ACTION act_Oper:
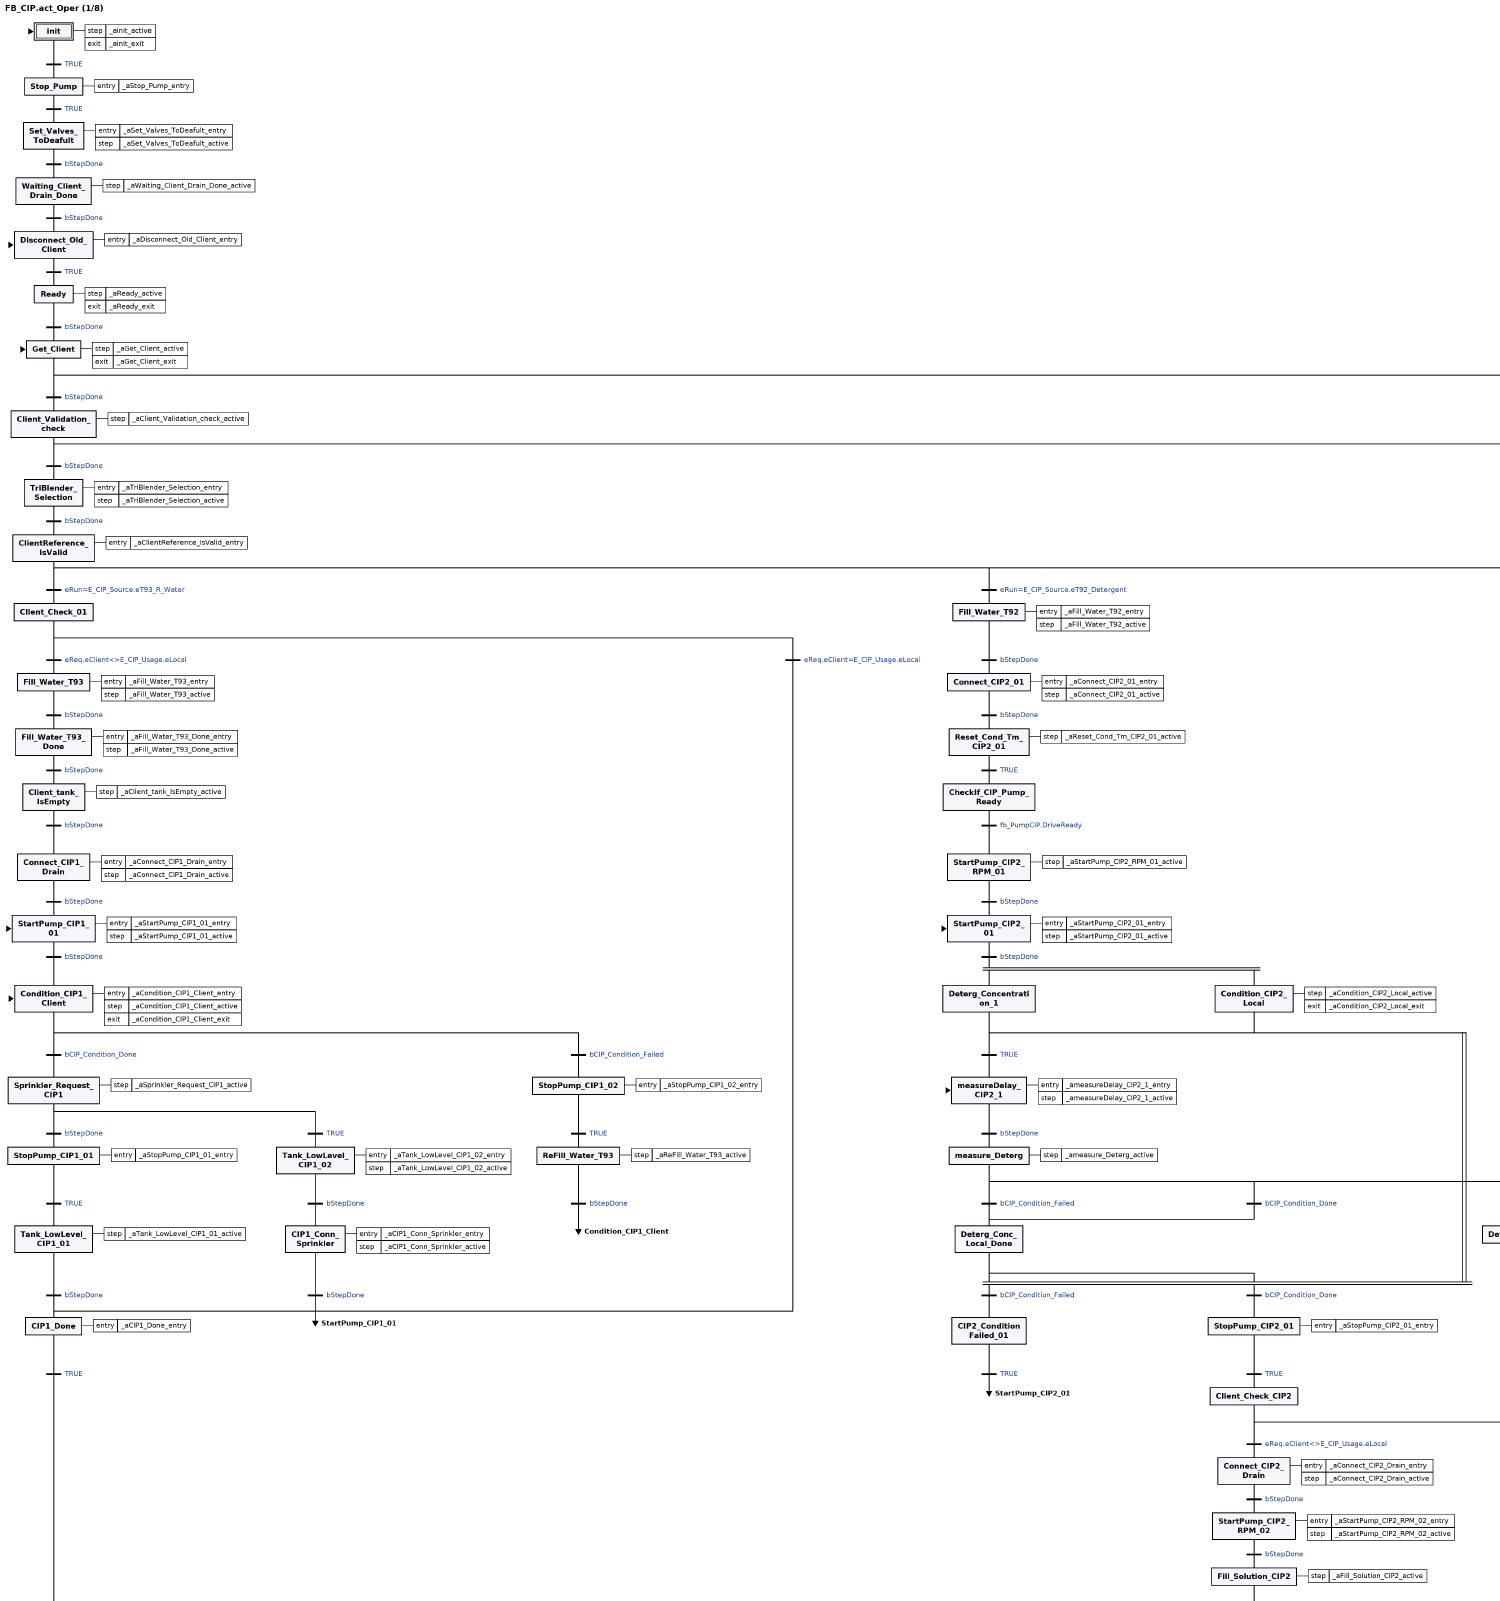
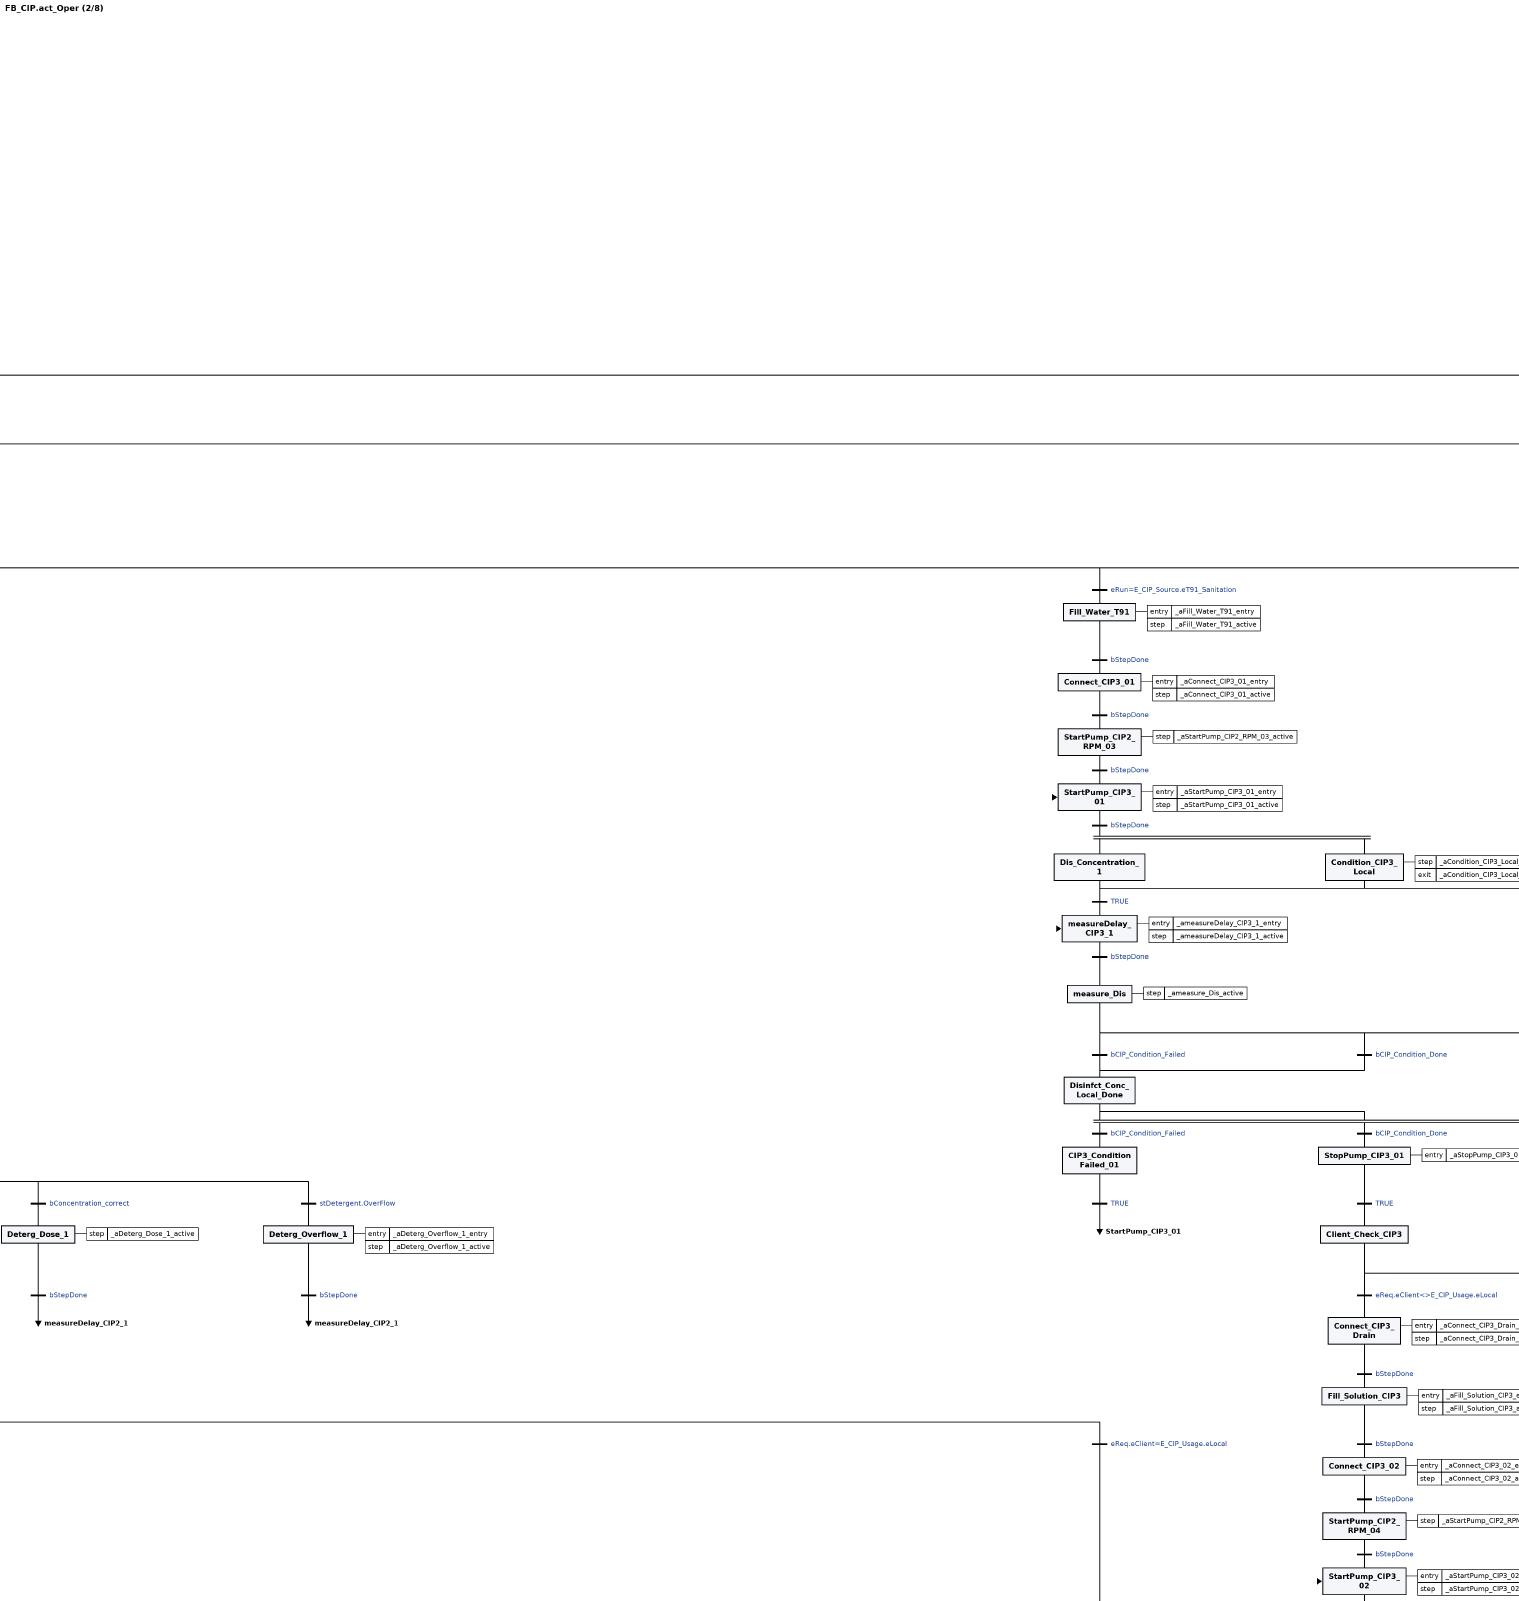
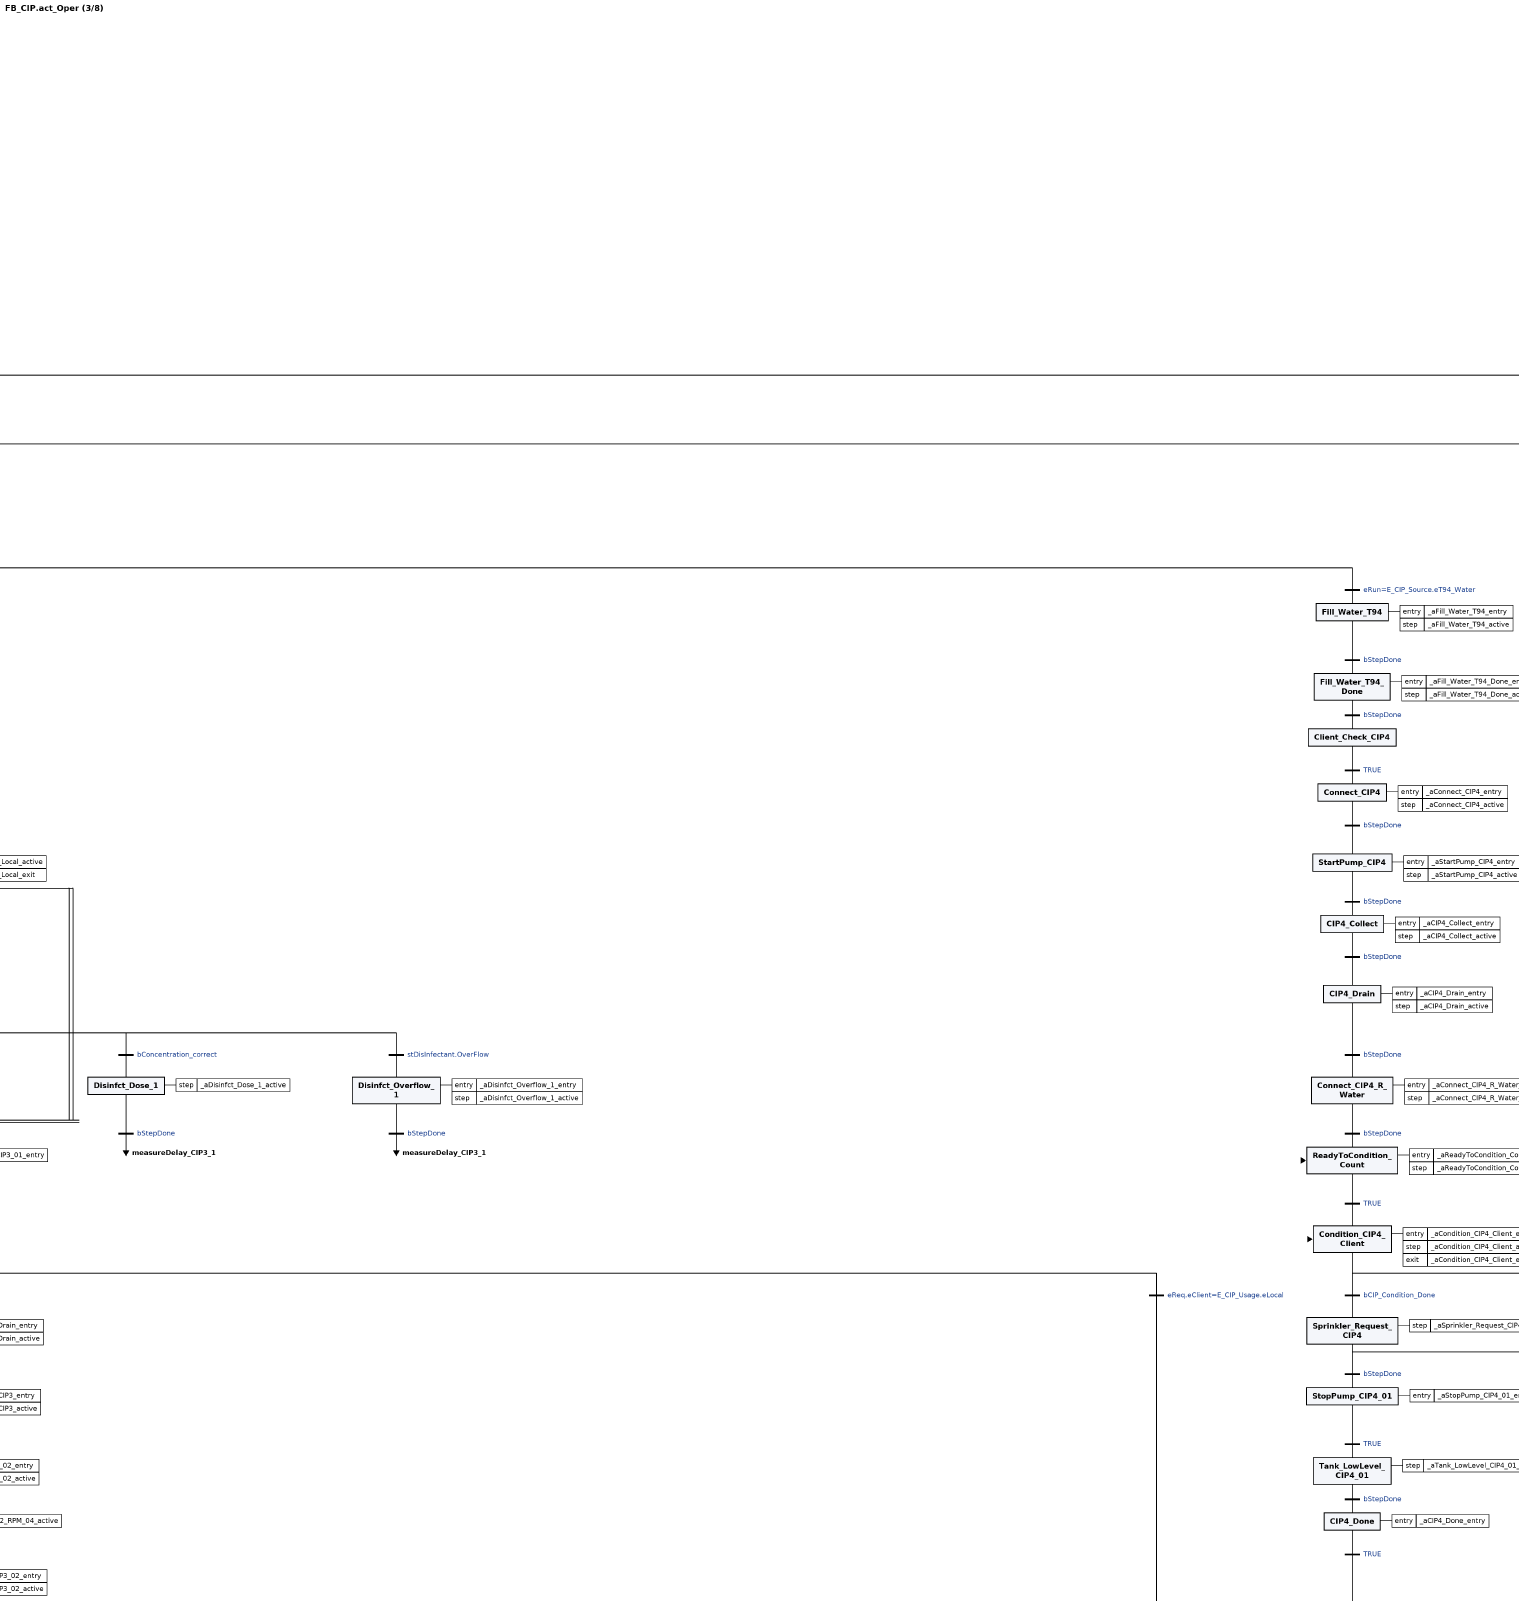
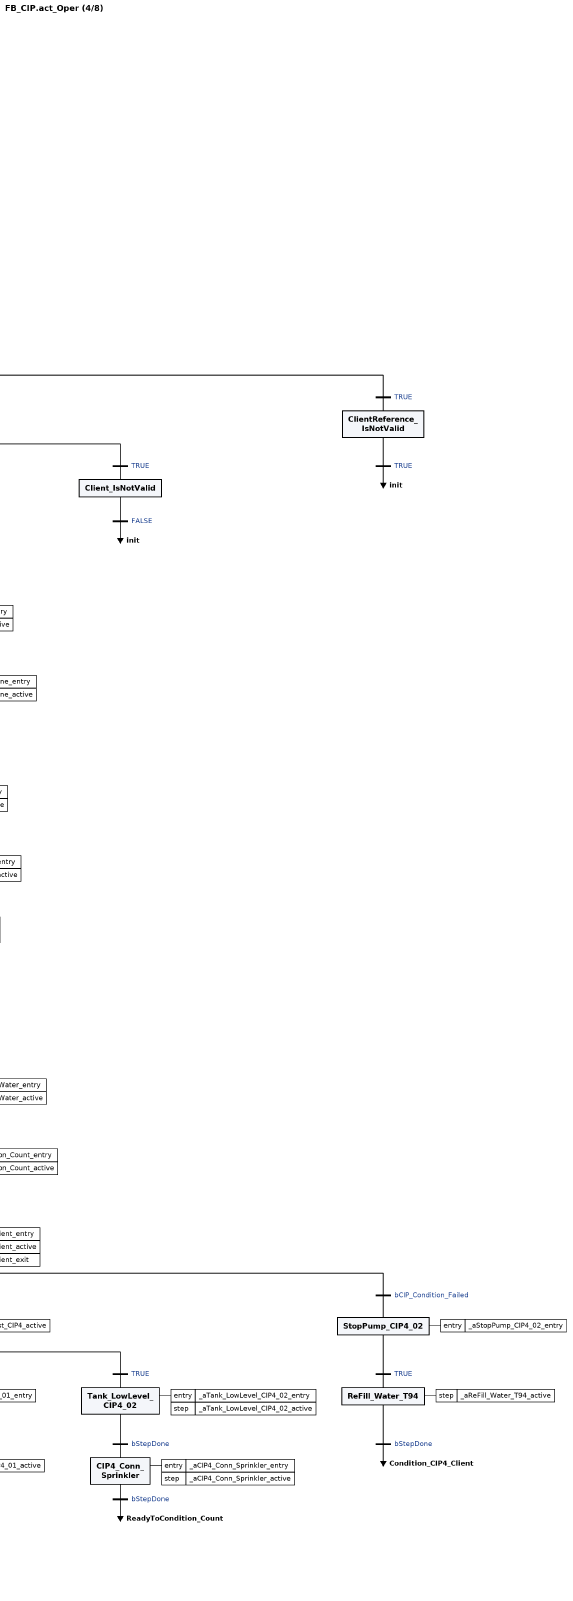
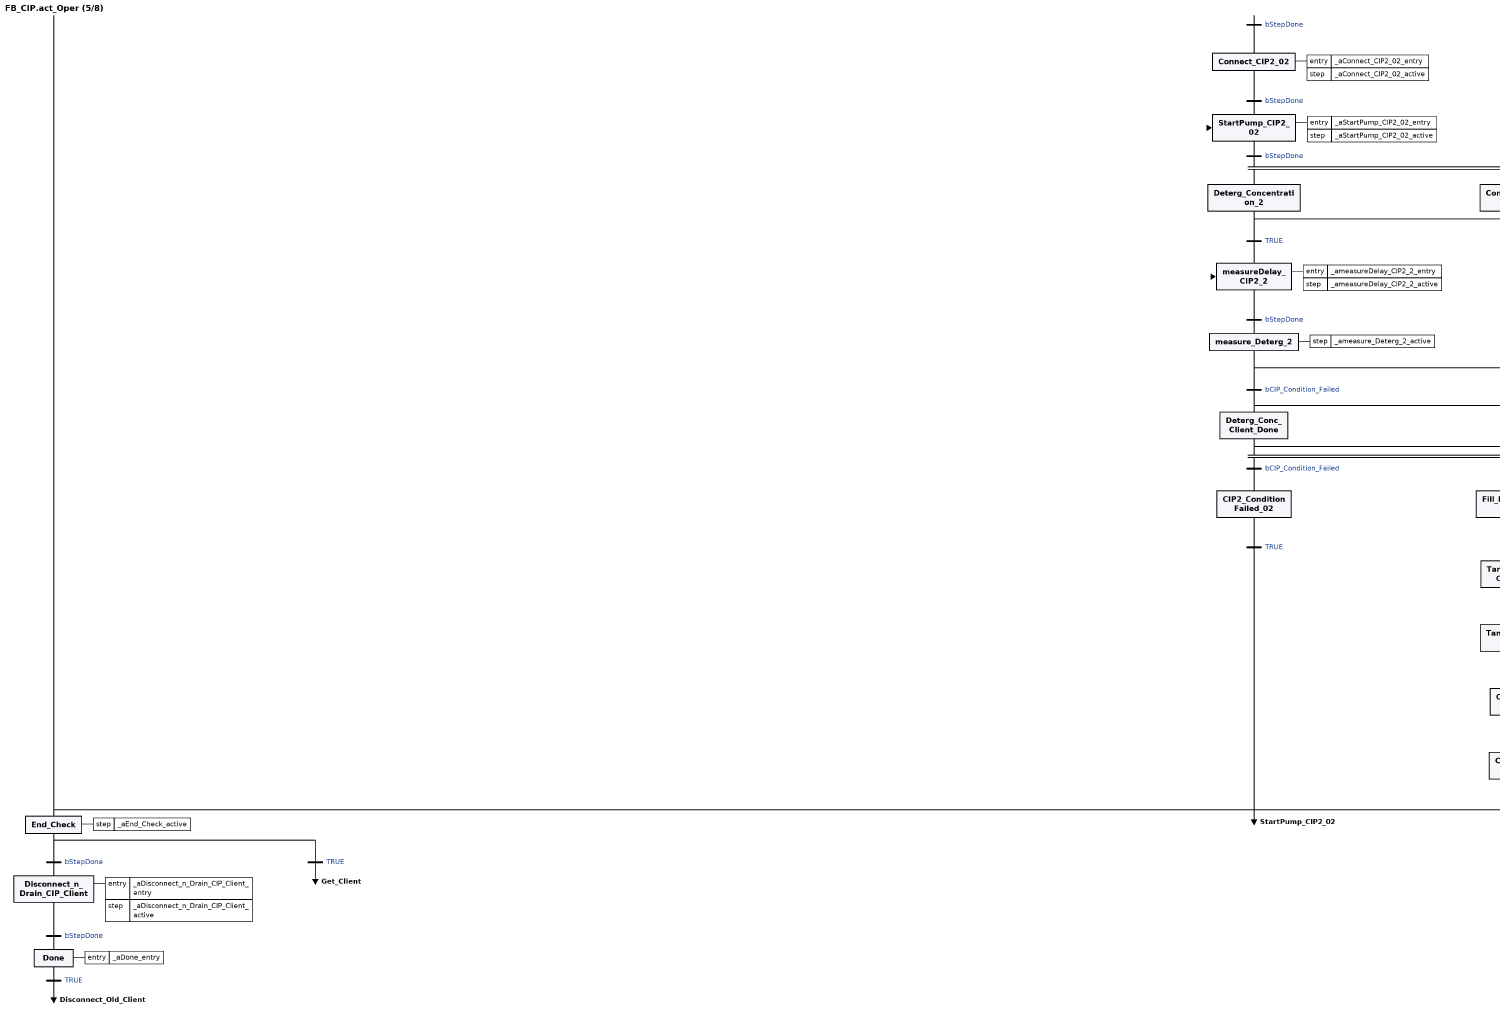
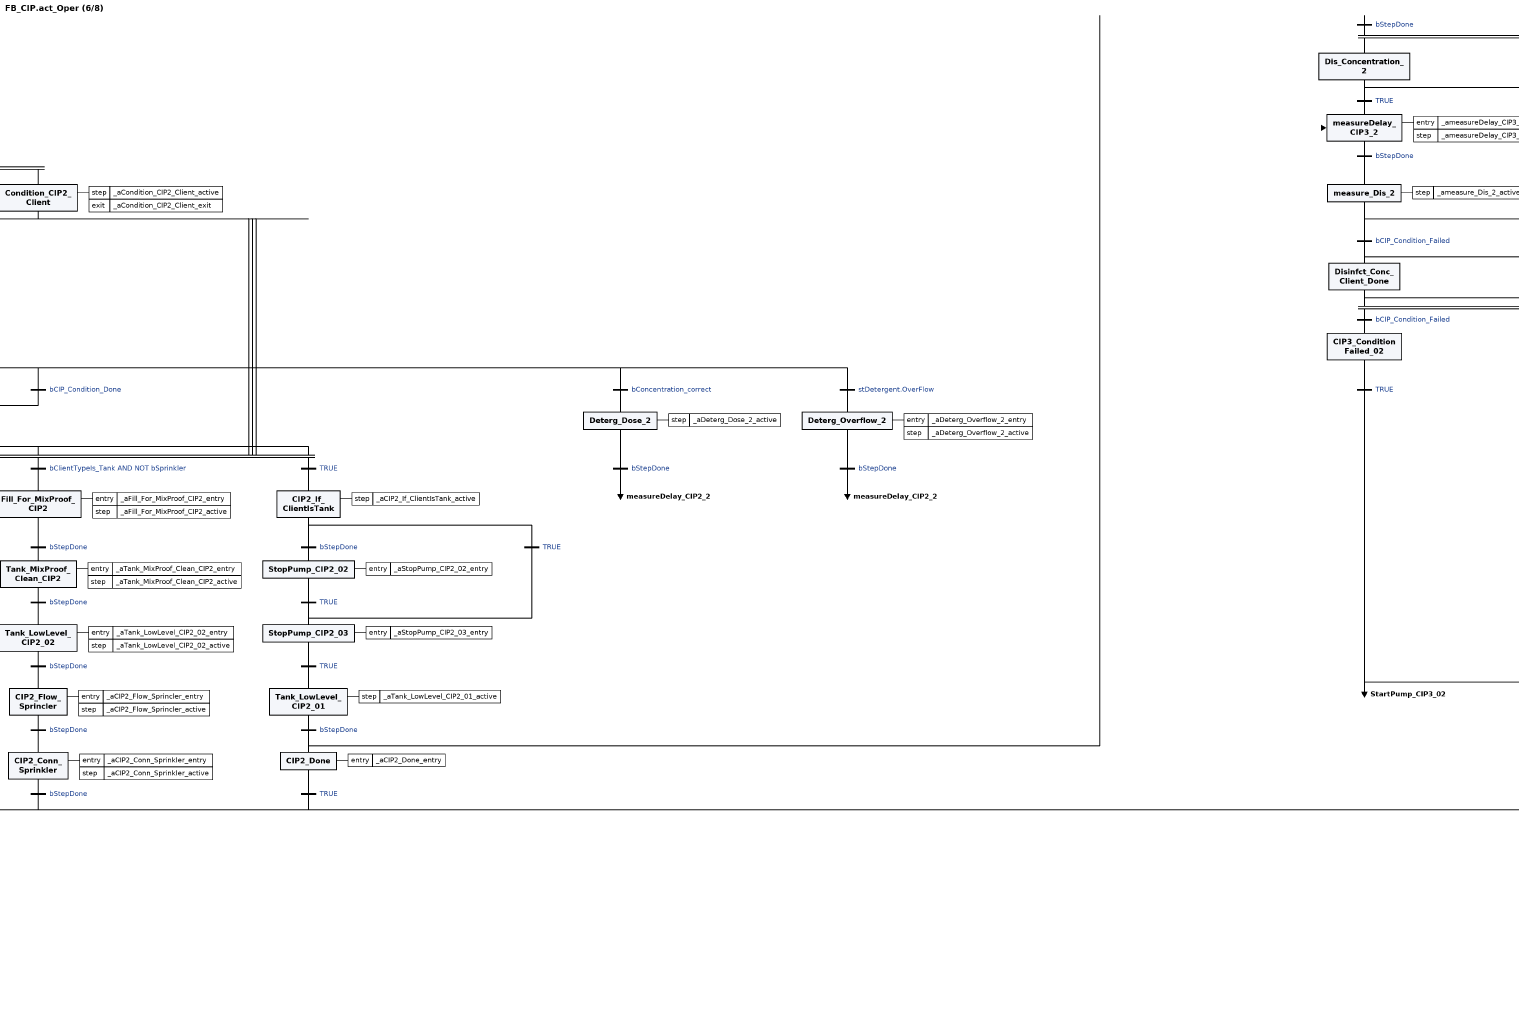
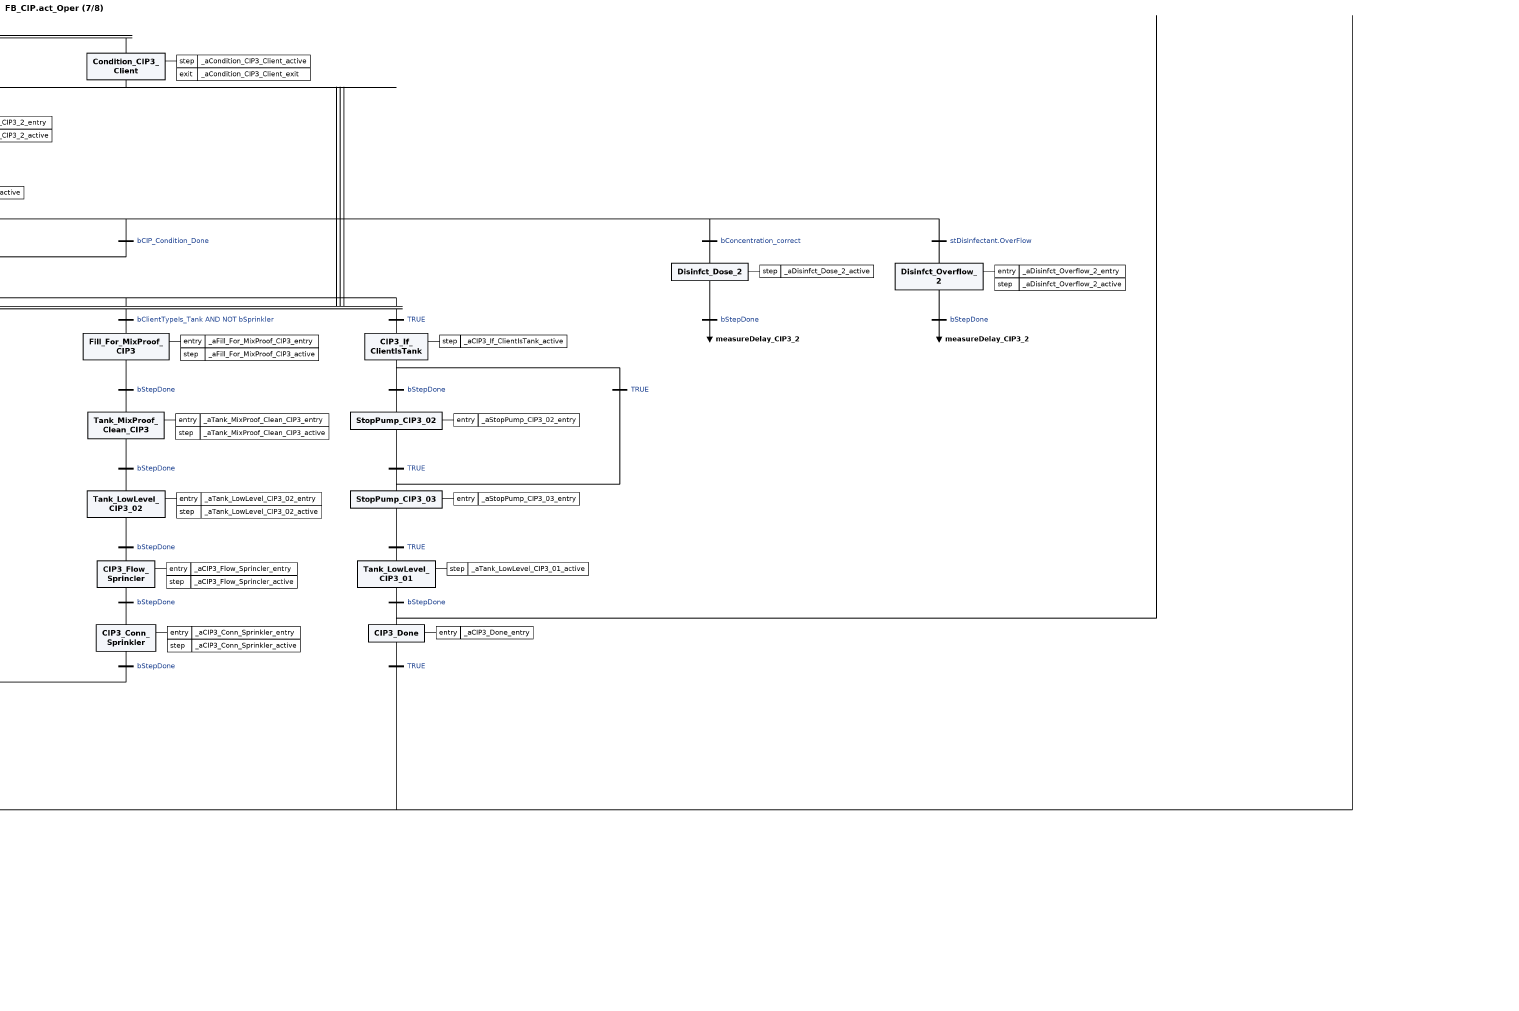
INITIAL_STEP init:
    _ainit_active(N);  // step action
    _ainit_exit(P0);  // exit action
END_STEP
TRANSITION FROM init TO Stop_Pump
    := TRUE;
END_TRANSITION
STEP Stop_Pump:
    _aStop_Pump_entry(P1);  // entry action
END_STEP
TRANSITION FROM Stop_Pump TO Set_Valves_ToDeafult
    := TRUE;
END_TRANSITION
STEP Set_Valves_ToDeafult:  // min time T#0.1s
    _aSet_Valves_ToDeafult_entry(P1);  // entry action
    _aSet_Valves_ToDeafult_active(N);  // step action
END_STEP
TRANSITION FROM Set_Valves_ToDeafult TO Waiting_Client_Drain_Done
    := bStepDone;
END_TRANSITION
STEP Waiting_Client_Drain_Done:  // min time T#0.1s
    _aWaiting_Client_Drain_Done_active(N);  // step action
END_STEP
TRANSITION FROM Waiting_Client_Drain_Done TO Disconnect_Old_Client
    := bStepDone;
END_TRANSITION
STEP Disconnect_Old_Client:
    _aDisconnect_Old_Client_entry(P1);  // entry action
END_STEP
TRANSITION FROM Disconnect_Old_Client TO Ready
    := TRUE;
END_TRANSITION
STEP Ready:
    _aReady_active(N);  // step action
    _aReady_exit(P0);  // exit action
END_STEP
TRANSITION FROM Ready TO Get_Client
    := bStepDone;
END_TRANSITION
STEP Get_Client:  // max time T#0.1s
    _aGet_Client_active(N);  // step action
    _aGet_Client_exit(P0);  // exit action
END_STEP
TRANSITION FROM Get_Client TO Client_Validation_check
    := bStepDone;
END_TRANSITION
TRANSITION FROM Get_Client TO ClientReference_IsNotValid
    := TRUE;
END_TRANSITION
STEP ClientReference_IsNotValid:  // min time T#2s
END_STEP
TRANSITION FROM ClientReference_IsNotValid TO init
    := TRUE;
END_TRANSITION
STEP Client_Validation_check:
    _aClient_Validation_check_active(N);  // step action
END_STEP
TRANSITION FROM Client_Validation_check TO TriBlender_Selection
    := bStepDone;
END_TRANSITION
STEP TriBlender_Selection:
    _aTriBlender_Selection_entry(P1);  // entry action
    _aTriBlender_Selection_active(N);  // step action
END_STEP
TRANSITION FROM TriBlender_Selection TO ClientReference_IsValid
    := bStepDone;
END_TRANSITION
TRANSITION FROM Client_Validation_check TO Client_IsNotValid
    := TRUE;
END_TRANSITION
STEP Client_IsNotValid:  // min time T#2s
END_STEP
TRANSITION FROM Client_IsNotValid TO init
    := FALSE;
END_TRANSITION
STEP ClientReference_IsValid:
    _aClientReference_IsValid_entry(P1);  // entry action
END_STEP
TRANSITION FROM ClientReference_IsValid TO Client_Check_01
    := eRun=E_CIP_Source.eT93_R_Water;
END_TRANSITION
// macro R_Water begins
STEP Client_Check_01:
END_STEP
TRANSITION FROM Client_Check_01 TO Fill_Water_T93
    := eReq.eClient<>E_CIP_Usage.eLocal;
END_TRANSITION
STEP Fill_Water_T93:
    _aFill_Water_T93_entry(P1);  // entry action
    _aFill_Water_T93_active(N);  // step action
END_STEP
TRANSITION FROM Fill_Water_T93 TO Fill_Water_T93_Done
    := bStepDone;
END_TRANSITION
STEP Fill_Water_T93_Done:
    _aFill_Water_T93_Done_entry(P1);  // entry action
    _aFill_Water_T93_Done_active(N);  // step action
END_STEP
TRANSITION FROM Fill_Water_T93_Done TO Client_tank_IsEmpty
    := bStepDone;
END_TRANSITION
STEP Client_tank_IsEmpty:  // min time T#5s
    _aClient_tank_IsEmpty_active(N);  // step action
END_STEP
TRANSITION FROM Client_tank_IsEmpty TO Connect_CIP1_Drain
    := bStepDone;
END_TRANSITION
STEP Connect_CIP1_Drain:
    _aConnect_CIP1_Drain_entry(P1);  // entry action
    _aConnect_CIP1_Drain_active(N);  // step action
END_STEP
TRANSITION FROM Connect_CIP1_Drain TO StartPump_CIP1_01
    := bStepDone;
END_TRANSITION
STEP StartPump_CIP1_01:
    _aStartPump_CIP1_01_entry(P1);  // entry action
    _aStartPump_CIP1_01_active(N);  // step action
END_STEP
TRANSITION FROM StartPump_CIP1_01 TO Condition_CIP1_Client
    := bStepDone;
END_TRANSITION
STEP Condition_CIP1_Client:
    _aCondition_CIP1_Client_entry(P1);  // entry action
    _aCondition_CIP1_Client_active(N);  // step action
    _aCondition_CIP1_Client_exit(P0);  // exit action
END_STEP
TRANSITION FROM Condition_CIP1_Client TO Sprinkler_Request_CIP1
    := bCIP_Condition_Done;
END_TRANSITION
STEP Sprinkler_Request_CIP1:
    _aSprinkler_Request_CIP1_active(N);  // step action
END_STEP
TRANSITION FROM Sprinkler_Request_CIP1 TO StopPump_CIP1_01
    := bStepDone;
END_TRANSITION
STEP StopPump_CIP1_01:
    _aStopPump_CIP1_01_entry(P1);  // entry action
END_STEP
TRANSITION FROM StopPump_CIP1_01 TO Tank_LowLevel_CIP1_01
    := TRUE;
END_TRANSITION
STEP Tank_LowLevel_CIP1_01:
    _aTank_LowLevel_CIP1_01_active(N);  // step action
END_STEP
TRANSITION FROM Tank_LowLevel_CIP1_01 TO CIP1_Done
    := bStepDone;
END_TRANSITION
TRANSITION FROM Sprinkler_Request_CIP1 TO Tank_LowLevel_CIP1_02
    := TRUE;
END_TRANSITION
STEP Tank_LowLevel_CIP1_02:
    _aTank_LowLevel_CIP1_02_entry(P1);  // entry action
    _aTank_LowLevel_CIP1_02_active(N);  // step action
END_STEP
TRANSITION FROM Tank_LowLevel_CIP1_02 TO CIP1_Conn_Sprinkler
    := bStepDone;
END_TRANSITION
STEP CIP1_Conn_Sprinkler:
    _aCIP1_Conn_Sprinkler_entry(P1);  // entry action
    _aCIP1_Conn_Sprinkler_active(N);  // step action
END_STEP
TRANSITION FROM CIP1_Conn_Sprinkler TO StartPump_CIP1_01
    := bStepDone;
END_TRANSITION
TRANSITION FROM Condition_CIP1_Client TO StopPump_CIP1_02
    := bCIP_Condition_Failed;
END_TRANSITION
STEP StopPump_CIP1_02:
    _aStopPump_CIP1_02_entry(P1);  // entry action
END_STEP
TRANSITION FROM StopPump_CIP1_02 TO ReFill_Water_T93
    := TRUE;
END_TRANSITION
STEP ReFill_Water_T93:
    _aReFill_Water_T93_active(N);  // step action
END_STEP
TRANSITION FROM ReFill_Water_T93 TO Condition_CIP1_Client
    := bStepDone;
END_TRANSITION
TRANSITION FROM Client_Check_01 TO CIP1_Done
    := eReq.eClient=E_CIP_Usage.eLocal;
END_TRANSITION
STEP CIP1_Done:  // min time T#2s
    _aCIP1_Done_entry(P1);  // entry action
END_STEP
TRANSITION FROM CIP1_Done TO End_Check
    := TRUE;
END_TRANSITION
TRANSITION FROM ClientReference_IsValid TO Fill_Water_T92
    := eRun=E_CIP_Source.eT92_Detergent;
END_TRANSITION
// macro Detergent begins
STEP Fill_Water_T92:
    _aFill_Water_T92_entry(P1);  // entry action
    _aFill_Water_T92_active(N);  // step action
END_STEP
TRANSITION FROM Fill_Water_T92 TO Connect_CIP2_01
    := bStepDone;
END_TRANSITION
STEP Connect_CIP2_01:
    _aConnect_CIP2_01_entry(P1);  // entry action
    _aConnect_CIP2_01_active(N);  // step action
END_STEP
TRANSITION FROM Connect_CIP2_01 TO Reset_Cond_Tm_CIP2_01
    := bStepDone;
END_TRANSITION
STEP Reset_Cond_Tm_CIP2_01:
    _aReset_Cond_Tm_CIP2_01_active(N);  // step action
END_STEP
TRANSITION FROM Reset_Cond_Tm_CIP2_01 TO CheckIf_CIP_Pump_Ready
    := TRUE;
END_TRANSITION
STEP CheckIf_CIP_Pump_Ready:
END_STEP
TRANSITION FROM CheckIf_CIP_Pump_Ready TO StartPump_CIP2_RPM_01
    := fb_PumpCIP.DriveReady;
END_TRANSITION
STEP StartPump_CIP2_RPM_01:
    _aStartPump_CIP2_RPM_01_active(N);  // step action
END_STEP
TRANSITION FROM StartPump_CIP2_RPM_01 TO StartPump_CIP2_01
    := bStepDone;
END_TRANSITION
STEP StartPump_CIP2_01:  // min time T#2s
    _aStartPump_CIP2_01_entry(P1);  // entry action
    _aStartPump_CIP2_01_active(N);  // step action
END_STEP
TRANSITION FROM StartPump_CIP2_01 TO (Deterg_Concentration_1, Condition_CIP2_Local)
    := bStepDone;
END_TRANSITION
STEP Deterg_Concentration_1:
END_STEP
TRANSITION FROM Deterg_Concentration_1 TO measureDelay_CIP2_1
    := TRUE;
END_TRANSITION
STEP measureDelay_CIP2_1:
    _ameasureDelay_CIP2_1_entry(P1);  // entry action
    _ameasureDelay_CIP2_1_active(N);  // step action
END_STEP
TRANSITION FROM measureDelay_CIP2_1 TO measure_Deterg
    := bStepDone;
END_TRANSITION
STEP measure_Deterg:  // min time t#1s
    _ameasure_Deterg_active(N);  // step action
END_STEP
TRANSITION FROM measure_Deterg TO Deterg_Conc_Local_Done
    := bCIP_Condition_Failed;
END_TRANSITION
TRANSITION FROM measure_Deterg TO Deterg_Conc_Local_Done
    := bCIP_Condition_Done;
END_TRANSITION
TRANSITION FROM measure_Deterg TO Deterg_Dose_1
    := bConcentration_correct;
END_TRANSITION
STEP Deterg_Dose_1:
    _aDeterg_Dose_1_active(N);  // step action
END_STEP
TRANSITION FROM Deterg_Dose_1 TO measureDelay_CIP2_1
    := bStepDone;
END_TRANSITION
TRANSITION FROM measure_Deterg TO Deterg_Overflow_1
    := stDetergent.OverFlow;
END_TRANSITION
STEP Deterg_Overflow_1:
    _aDeterg_Overflow_1_entry(P1);  // entry action
    _aDeterg_Overflow_1_active(N);  // step action
END_STEP
TRANSITION FROM Deterg_Overflow_1 TO measureDelay_CIP2_1
    := bStepDone;
END_TRANSITION
STEP Deterg_Conc_Local_Done:
END_STEP
STEP Condition_CIP2_Local:
    _aCondition_CIP2_Local_active(N);  // step action
    _aCondition_CIP2_Local_exit(P0);  // exit action
END_STEP
TRANSITION FROM (Deterg_Conc_Local_Done, Condition_CIP2_Local) TO CIP2_ConditionFailed_01
    := bCIP_Condition_Failed;
END_TRANSITION
STEP CIP2_ConditionFailed_01:
END_STEP
TRANSITION FROM CIP2_ConditionFailed_01 TO StartPump_CIP2_01
    := TRUE;
END_TRANSITION
TRANSITION FROM (Deterg_Conc_Local_Done, Condition_CIP2_Local) TO StopPump_CIP2_01
    := bCIP_Condition_Done;
END_TRANSITION
STEP StopPump_CIP2_01:
    _aStopPump_CIP2_01_entry(P1);  // entry action
END_STEP
TRANSITION FROM StopPump_CIP2_01 TO Client_Check_CIP2
    := TRUE;
END_TRANSITION
STEP Client_Check_CIP2:
END_STEP
TRANSITION FROM Client_Check_CIP2 TO Connect_CIP2_Drain
    := eReq.eClient<>E_CIP_Usage.eLocal;
END_TRANSITION
STEP Connect_CIP2_Drain:
    _aConnect_CIP2_Drain_entry(P1);  // entry action
    _aConnect_CIP2_Drain_active(N);  // step action
END_STEP
TRANSITION FROM Connect_CIP2_Drain TO StartPump_CIP2_RPM_02
    := bStepDone;
END_TRANSITION
STEP StartPump_CIP2_RPM_02:
    _aStartPump_CIP2_RPM_02_entry(P1);  // entry action
    _aStartPump_CIP2_RPM_02_active(N);  // step action
END_STEP
TRANSITION FROM StartPump_CIP2_RPM_02 TO Fill_Solution_CIP2
    := bStepDone;
END_TRANSITION
STEP Fill_Solution_CIP2:
    _aFill_Solution_CIP2_active(N);  // step action
END_STEP
TRANSITION FROM Fill_Solution_CIP2 TO Connect_CIP2_02
    := bStepDone;
END_TRANSITION
STEP Connect_CIP2_02:
    _aConnect_CIP2_02_entry(P1);  // entry action
    _aConnect_CIP2_02_active(N);  // step action
END_STEP
TRANSITION FROM Connect_CIP2_02 TO StartPump_CIP2_02
    := bStepDone;
END_TRANSITION
STEP StartPump_CIP2_02:  // min time T#2s
    _aStartPump_CIP2_02_entry(P1);  // entry action
    _aStartPump_CIP2_02_active(N);  // step action
END_STEP
TRANSITION FROM StartPump_CIP2_02 TO (Deterg_Concentration_2, Condition_CIP2_Client)
    := bStepDone;
END_TRANSITION
STEP Deterg_Concentration_2:
END_STEP
TRANSITION FROM Deterg_Concentration_2 TO measureDelay_CIP2_2
    := TRUE;
END_TRANSITION
STEP measureDelay_CIP2_2:
    _ameasureDelay_CIP2_2_entry(P1);  // entry action
    _ameasureDelay_CIP2_2_active(N);  // step action
END_STEP
TRANSITION FROM measureDelay_CIP2_2 TO measure_Deterg_2
    := bStepDone;
END_TRANSITION
STEP measure_Deterg_2:  // min time t#1s
    _ameasure_Deterg_2_active(N);  // step action
END_STEP
TRANSITION FROM measure_Deterg_2 TO Deterg_Conc_Client_Done
    := bCIP_Condition_Failed;
END_TRANSITION
TRANSITION FROM measure_Deterg_2 TO Deterg_Conc_Client_Done
    := bCIP_Condition_Done;
END_TRANSITION
TRANSITION FROM measure_Deterg_2 TO Deterg_Dose_2
    := bConcentration_correct;
END_TRANSITION
STEP Deterg_Dose_2:
    _aDeterg_Dose_2_active(N);  // step action
END_STEP
TRANSITION FROM Deterg_Dose_2 TO measureDelay_CIP2_2
    := bStepDone;
END_TRANSITION
TRANSITION FROM measure_Deterg_2 TO Deterg_Overflow_2
    := stDetergent.OverFlow;
END_TRANSITION
STEP Deterg_Overflow_2:
    _aDeterg_Overflow_2_entry(P1);  // entry action
    _aDeterg_Overflow_2_active(N);  // step action
END_STEP
TRANSITION FROM Deterg_Overflow_2 TO measureDelay_CIP2_2
    := bStepDone;
END_TRANSITION
STEP Deterg_Conc_Client_Done:
END_STEP
STEP Condition_CIP2_Client:
    _aCondition_CIP2_Client_active(N);  // step action
    _aCondition_CIP2_Client_exit(P0);  // exit action
END_STEP
TRANSITION FROM (Deterg_Conc_Client_Done, Condition_CIP2_Client) TO CIP2_ConditionFailed_02
    := bCIP_Condition_Failed;
END_TRANSITION
STEP CIP2_ConditionFailed_02:
END_STEP
TRANSITION FROM CIP2_ConditionFailed_02 TO StartPump_CIP2_02
    := TRUE;
END_TRANSITION
TRANSITION FROM (Deterg_Conc_Client_Done, Condition_CIP2_Client) TO Fill_For_MixProof_CIP2
    := bClientTypeIs_Tank AND NOT bSprinkler;
END_TRANSITION
STEP Fill_For_MixProof_CIP2:
    _aFill_For_MixProof_CIP2_entry(P1);  // entry action
    _aFill_For_MixProof_CIP2_active(N);  // step action
END_STEP
TRANSITION FROM Fill_For_MixProof_CIP2 TO Tank_MixProof_Clean_CIP2
    := bStepDone;
END_TRANSITION
STEP Tank_MixProof_Clean_CIP2:
    _aTank_MixProof_Clean_CIP2_entry(P1);  // entry action
    _aTank_MixProof_Clean_CIP2_active(N);  // step action
END_STEP
TRANSITION FROM Tank_MixProof_Clean_CIP2 TO Tank_LowLevel_CIP2_02
    := bStepDone;
END_TRANSITION
STEP Tank_LowLevel_CIP2_02:
    _aTank_LowLevel_CIP2_02_entry(P1);  // entry action
    _aTank_LowLevel_CIP2_02_active(N);  // step action
END_STEP
TRANSITION FROM Tank_LowLevel_CIP2_02 TO CIP2_Flow_Sprincler
    := bStepDone;
END_TRANSITION
STEP CIP2_Flow_Sprincler:
    _aCIP2_Flow_Sprincler_entry(P1);  // entry action
    _aCIP2_Flow_Sprincler_active(N);  // step action
END_STEP
TRANSITION FROM CIP2_Flow_Sprincler TO CIP2_Conn_Sprinkler
    := bStepDone;
END_TRANSITION
STEP CIP2_Conn_Sprinkler:
    _aCIP2_Conn_Sprinkler_entry(P1);  // entry action
    _aCIP2_Conn_Sprinkler_active(N);  // step action
END_STEP
TRANSITION FROM CIP2_Conn_Sprinkler TO StartPump_CIP2_02
    := bStepDone;
END_TRANSITION
TRANSITION FROM (Deterg_Conc_Client_Done, Condition_CIP2_Client) TO CIP2_If_ClientIsTank
    := TRUE;
END_TRANSITION
STEP CIP2_If_ClientIsTank:
    _aCIP2_If_ClientIsTank_active(N);  // step action
END_STEP
TRANSITION FROM CIP2_If_ClientIsTank TO StopPump_CIP2_02
    := bStepDone;
END_TRANSITION
STEP StopPump_CIP2_02:
    _aStopPump_CIP2_02_entry(P1);  // entry action
END_STEP
TRANSITION FROM StopPump_CIP2_02 TO StopPump_CIP2_03
    := TRUE;
END_TRANSITION
TRANSITION FROM CIP2_If_ClientIsTank TO StopPump_CIP2_03
    := TRUE;
END_TRANSITION
STEP StopPump_CIP2_03:
    _aStopPump_CIP2_03_entry(P1);  // entry action
END_STEP
TRANSITION FROM StopPump_CIP2_03 TO Tank_LowLevel_CIP2_01
    := TRUE;
END_TRANSITION
STEP Tank_LowLevel_CIP2_01:
    _aTank_LowLevel_CIP2_01_active(N);  // step action
END_STEP
TRANSITION FROM Tank_LowLevel_CIP2_01 TO CIP2_Done
    := bStepDone;
END_TRANSITION
TRANSITION FROM Client_Check_CIP2 TO CIP2_Done
    := eReq.eClient=E_CIP_Usage.eLocal;
END_TRANSITION
STEP CIP2_Done:  // min time T#2s
    _aCIP2_Done_entry(P1);  // entry action
END_STEP
TRANSITION FROM CIP2_Done TO End_Check
    := TRUE;
END_TRANSITION
TRANSITION FROM ClientReference_IsValid TO Fill_Water_T91
    := eRun=E_CIP_Source.eT91_Sanitation;
END_TRANSITION
// macro DisInfection begins
STEP Fill_Water_T91:
    _aFill_Water_T91_entry(P1);  // entry action
    _aFill_Water_T91_active(N);  // step action
END_STEP
TRANSITION FROM Fill_Water_T91 TO Connect_CIP3_01
    := bStepDone;
END_TRANSITION
STEP Connect_CIP3_01:
    _aConnect_CIP3_01_entry(P1);  // entry action
    _aConnect_CIP3_01_active(N);  // step action
END_STEP
TRANSITION FROM Connect_CIP3_01 TO StartPump_CIP2_RPM_03
    := bStepDone;
END_TRANSITION
STEP StartPump_CIP2_RPM_03:
    _aStartPump_CIP2_RPM_03_active(N);  // step action
END_STEP
TRANSITION FROM StartPump_CIP2_RPM_03 TO StartPump_CIP3_01
    := bStepDone;
END_TRANSITION
STEP StartPump_CIP3_01:  // min time T#3s
    _aStartPump_CIP3_01_entry(P1);  // entry action
    _aStartPump_CIP3_01_active(N);  // step action
END_STEP
TRANSITION FROM StartPump_CIP3_01 TO (Dis_Concentration_1, Condition_CIP3_Local)
    := bStepDone;
END_TRANSITION
STEP Dis_Concentration_1:
END_STEP
TRANSITION FROM Dis_Concentration_1 TO measureDelay_CIP3_1
    := TRUE;
END_TRANSITION
STEP measureDelay_CIP3_1:
    _ameasureDelay_CIP3_1_entry(P1);  // entry action
    _ameasureDelay_CIP3_1_active(N);  // step action
END_STEP
TRANSITION FROM measureDelay_CIP3_1 TO measure_Dis
    := bStepDone;
END_TRANSITION
STEP measure_Dis:  // min time t#1s
    _ameasure_Dis_active(N);  // step action
END_STEP
TRANSITION FROM measure_Dis TO Disinfct_Conc_Local_Done
    := bCIP_Condition_Failed;
END_TRANSITION
TRANSITION FROM measure_Dis TO Disinfct_Conc_Local_Done
    := bCIP_Condition_Done;
END_TRANSITION
TRANSITION FROM measure_Dis TO Disinfct_Dose_1
    := bConcentration_correct;
END_TRANSITION
STEP Disinfct_Dose_1:
    _aDisinfct_Dose_1_active(N);  // step action
END_STEP
TRANSITION FROM Disinfct_Dose_1 TO measureDelay_CIP3_1
    := bStepDone;
END_TRANSITION
TRANSITION FROM measure_Dis TO Disinfct_Overflow_1
    := stDisInfectant.OverFlow;
END_TRANSITION
STEP Disinfct_Overflow_1:
    _aDisinfct_Overflow_1_entry(P1);  // entry action
    _aDisinfct_Overflow_1_active(N);  // step action
END_STEP
TRANSITION FROM Disinfct_Overflow_1 TO measureDelay_CIP3_1
    := bStepDone;
END_TRANSITION
STEP Disinfct_Conc_Local_Done:
END_STEP
STEP Condition_CIP3_Local:
    _aCondition_CIP3_Local_active(N);  // step action
    _aCondition_CIP3_Local_exit(P0);  // exit action
END_STEP
TRANSITION FROM (Disinfct_Conc_Local_Done, Condition_CIP3_Local) TO CIP3_ConditionFailed_01
    := bCIP_Condition_Failed;
END_TRANSITION
STEP CIP3_ConditionFailed_01:
END_STEP
TRANSITION FROM CIP3_ConditionFailed_01 TO StartPump_CIP3_01
    := TRUE;
END_TRANSITION
TRANSITION FROM (Disinfct_Conc_Local_Done, Condition_CIP3_Local) TO StopPump_CIP3_01
    := bCIP_Condition_Done;
END_TRANSITION
STEP StopPump_CIP3_01:  // min time T#5s
    _aStopPump_CIP3_01_entry(P1);  // entry action
END_STEP
TRANSITION FROM StopPump_CIP3_01 TO Client_Check_CIP3
    := TRUE;
END_TRANSITION
STEP Client_Check_CIP3:
END_STEP
TRANSITION FROM Client_Check_CIP3 TO Connect_CIP3_Drain
    := eReq.eClient<>E_CIP_Usage.eLocal;
END_TRANSITION
STEP Connect_CIP3_Drain:
    _aConnect_CIP3_Drain_entry(P1);  // entry action
    _aConnect_CIP3_Drain_active(N);  // step action
END_STEP
TRANSITION FROM Connect_CIP3_Drain TO Fill_Solution_CIP3
    := bStepDone;
END_TRANSITION
STEP Fill_Solution_CIP3:
    _aFill_Solution_CIP3_entry(P1);  // entry action
    _aFill_Solution_CIP3_active(N);  // step action
END_STEP
TRANSITION FROM Fill_Solution_CIP3 TO Connect_CIP3_02
    := bStepDone;
END_TRANSITION
STEP Connect_CIP3_02:
    _aConnect_CIP3_02_entry(P1);  // entry action
    _aConnect_CIP3_02_active(N);  // step action
END_STEP
TRANSITION FROM Connect_CIP3_02 TO StartPump_CIP2_RPM_04
    := bStepDone;
END_TRANSITION
STEP StartPump_CIP2_RPM_04:
    _aStartPump_CIP2_RPM_04_active(N);  // step action
END_STEP
TRANSITION FROM StartPump_CIP2_RPM_04 TO StartPump_CIP3_02
    := bStepDone;
END_TRANSITION
STEP StartPump_CIP3_02:  // min time T#1s
    _aStartPump_CIP3_02_entry(P1);  // entry action
    _aStartPump_CIP3_02_active(N);  // step action
END_STEP
TRANSITION FROM StartPump_CIP3_02 TO (Dis_Concentration_2, Condition_CIP3_Client)
    := bStepDone;
END_TRANSITION
STEP Dis_Concentration_2:
END_STEP
TRANSITION FROM Dis_Concentration_2 TO measureDelay_CIP3_2
    := TRUE;
END_TRANSITION
STEP measureDelay_CIP3_2:
    _ameasureDelay_CIP3_2_entry(P1);  // entry action
    _ameasureDelay_CIP3_2_active(N);  // step action
END_STEP
TRANSITION FROM measureDelay_CIP3_2 TO measure_Dis_2
    := bStepDone;
END_TRANSITION
STEP measure_Dis_2:  // min time t#1s
    _ameasure_Dis_2_active(N);  // step action
END_STEP
TRANSITION FROM measure_Dis_2 TO Disinfct_Conc_Client_Done
    := bCIP_Condition_Failed;
END_TRANSITION
TRANSITION FROM measure_Dis_2 TO Disinfct_Conc_Client_Done
    := bCIP_Condition_Done;
END_TRANSITION
TRANSITION FROM measure_Dis_2 TO Disinfct_Dose_2
    := bConcentration_correct;
END_TRANSITION
STEP Disinfct_Dose_2:
    _aDisinfct_Dose_2_active(N);  // step action
END_STEP
TRANSITION FROM Disinfct_Dose_2 TO measureDelay_CIP3_2
    := bStepDone;
END_TRANSITION
TRANSITION FROM measure_Dis_2 TO Disinfct_Overflow_2
    := stDisInfectant.OverFlow;
END_TRANSITION
STEP Disinfct_Overflow_2:
    _aDisinfct_Overflow_2_entry(P1);  // entry action
    _aDisinfct_Overflow_2_active(N);  // step action
END_STEP
TRANSITION FROM Disinfct_Overflow_2 TO measureDelay_CIP3_2
    := bStepDone;
END_TRANSITION
STEP Disinfct_Conc_Client_Done:
END_STEP
STEP Condition_CIP3_Client:
    _aCondition_CIP3_Client_active(N);  // step action
    _aCondition_CIP3_Client_exit(P0);  // exit action
END_STEP
TRANSITION FROM (Disinfct_Conc_Client_Done, Condition_CIP3_Client) TO CIP3_ConditionFailed_02
    := bCIP_Condition_Failed;
END_TRANSITION
STEP CIP3_ConditionFailed_02:
END_STEP
TRANSITION FROM CIP3_ConditionFailed_02 TO StartPump_CIP3_02
    := TRUE;
END_TRANSITION
TRANSITION FROM (Disinfct_Conc_Client_Done, Condition_CIP3_Client) TO Fill_For_MixProof_CIP3
    := bClientTypeIs_Tank AND NOT bSprinkler;
END_TRANSITION
STEP Fill_For_MixProof_CIP3:
    _aFill_For_MixProof_CIP3_entry(P1);  // entry action
    _aFill_For_MixProof_CIP3_active(N);  // step action
END_STEP
TRANSITION FROM Fill_For_MixProof_CIP3 TO Tank_MixProof_Clean_CIP3
    := bStepDone;
END_TRANSITION
STEP Tank_MixProof_Clean_CIP3:
    _aTank_MixProof_Clean_CIP3_entry(P1);  // entry action
    _aTank_MixProof_Clean_CIP3_active(N);  // step action
END_STEP
TRANSITION FROM Tank_MixProof_Clean_CIP3 TO Tank_LowLevel_CIP3_02
    := bStepDone;
END_TRANSITION
STEP Tank_LowLevel_CIP3_02:
    _aTank_LowLevel_CIP3_02_entry(P1);  // entry action
    _aTank_LowLevel_CIP3_02_active(N);  // step action
END_STEP
TRANSITION FROM Tank_LowLevel_CIP3_02 TO CIP3_Flow_Sprincler
    := bStepDone;
END_TRANSITION
STEP CIP3_Flow_Sprincler:
    _aCIP3_Flow_Sprincler_entry(P1);  // entry action
    _aCIP3_Flow_Sprincler_active(N);  // step action
END_STEP
TRANSITION FROM CIP3_Flow_Sprincler TO CIP3_Conn_Sprinkler
    := bStepDone;
END_TRANSITION
STEP CIP3_Conn_Sprinkler:
    _aCIP3_Conn_Sprinkler_entry(P1);  // entry action
    _aCIP3_Conn_Sprinkler_active(N);  // step action
END_STEP
TRANSITION FROM CIP3_Conn_Sprinkler TO StartPump_CIP3_02
    := bStepDone;
END_TRANSITION
TRANSITION FROM (Disinfct_Conc_Client_Done, Condition_CIP3_Client) TO CIP3_If_ClientIsTank
    := TRUE;
END_TRANSITION
STEP CIP3_If_ClientIsTank:
    _aCIP3_If_ClientIsTank_active(N);  // step action
END_STEP
TRANSITION FROM CIP3_If_ClientIsTank TO StopPump_CIP3_02
    := bStepDone;
END_TRANSITION
STEP StopPump_CIP3_02:  // min time T#2s
    _aStopPump_CIP3_02_entry(P1);  // entry action
END_STEP
TRANSITION FROM StopPump_CIP3_02 TO StopPump_CIP3_03
    := TRUE;
END_TRANSITION
TRANSITION FROM CIP3_If_ClientIsTank TO StopPump_CIP3_03
    := TRUE;
END_TRANSITION
STEP StopPump_CIP3_03:
    _aStopPump_CIP3_03_entry(P1);  // entry action
END_STEP
TRANSITION FROM StopPump_CIP3_03 TO Tank_LowLevel_CIP3_01
    := TRUE;
END_TRANSITION
STEP Tank_LowLevel_CIP3_01:
    _aTank_LowLevel_CIP3_01_active(N);  // step action
END_STEP
TRANSITION FROM Tank_LowLevel_CIP3_01 TO CIP3_Done
    := bStepDone;
END_TRANSITION
TRANSITION FROM Client_Check_CIP3 TO CIP3_Done
    := eReq.eClient=E_CIP_Usage.eLocal;
END_TRANSITION
STEP CIP3_Done:  // min time T#2s
    _aCIP3_Done_entry(P1);  // entry action
END_STEP
TRANSITION FROM CIP3_Done TO End_Check
    := TRUE;
END_TRANSITION
TRANSITION FROM ClientReference_IsValid TO Fill_Water_T94
    := eRun=E_CIP_Source.eT94_Water;
END_TRANSITION
// macro Water begins
STEP Fill_Water_T94:
    _aFill_Water_T94_entry(P1);  // entry action
    _aFill_Water_T94_active(N);  // step action
END_STEP
TRANSITION FROM Fill_Water_T94 TO Fill_Water_T94_Done
    := bStepDone;
END_TRANSITION
STEP Fill_Water_T94_Done:
    _aFill_Water_T94_Done_entry(P1);  // entry action
    _aFill_Water_T94_Done_active(N);  // step action
END_STEP
TRANSITION FROM Fill_Water_T94_Done TO Client_Check_CIP4
    := bStepDone;
END_TRANSITION
STEP Client_Check_CIP4:
END_STEP
TRANSITION FROM Client_Check_CIP4 TO Connect_CIP4
    := TRUE;
END_TRANSITION
STEP Connect_CIP4:
    _aConnect_CIP4_entry(P1);  // entry action
    _aConnect_CIP4_active(N);  // step action
END_STEP
TRANSITION FROM Connect_CIP4 TO StartPump_CIP4
    := bStepDone;
END_TRANSITION
STEP StartPump_CIP4:  // min time T#3s
    _aStartPump_CIP4_entry(P1);  // entry action
    _aStartPump_CIP4_active(N);  // step action
END_STEP
TRANSITION FROM StartPump_CIP4 TO CIP4_Collect
    := bStepDone;
END_TRANSITION
STEP CIP4_Collect:  // min time T#5s
    _aCIP4_Collect_entry(P1);  // entry action
    _aCIP4_Collect_active(N);  // step action
END_STEP
TRANSITION FROM CIP4_Collect TO CIP4_Drain
    := bStepDone;
END_TRANSITION
STEP CIP4_Drain:  // min time T#5s
    _aCIP4_Drain_entry(P1);  // entry action
    _aCIP4_Drain_active(N);  // step action
END_STEP
TRANSITION FROM CIP4_Drain TO Connect_CIP4_R_Water
    := bStepDone;
END_TRANSITION
STEP Connect_CIP4_R_Water:  // min time T#5s
    _aConnect_CIP4_R_Water_entry(P1);  // entry action
    _aConnect_CIP4_R_Water_active(N);  // step action
END_STEP
TRANSITION FROM Connect_CIP4_R_Water TO ReadyToCondition_Count
    := bStepDone;
END_TRANSITION
STEP ReadyToCondition_Count:
    _aReadyToCondition_Count_entry(P1);  // entry action
    _aReadyToCondition_Count_active(N);  // step action
END_STEP
TRANSITION FROM ReadyToCondition_Count TO Condition_CIP4_Client
    := TRUE;
END_TRANSITION
STEP Condition_CIP4_Client:
    _aCondition_CIP4_Client_entry(P1);  // entry action
    _aCondition_CIP4_Client_active(N);  // step action
    _aCondition_CIP4_Client_exit(P0);  // exit action
END_STEP
TRANSITION FROM Condition_CIP4_Client TO Sprinkler_Request_CIP4
    := bCIP_Condition_Done;
END_TRANSITION
STEP Sprinkler_Request_CIP4:
    _aSprinkler_Request_CIP4_active(N);  // step action
END_STEP
TRANSITION FROM Sprinkler_Request_CIP4 TO StopPump_CIP4_01
    := bStepDone;
END_TRANSITION
STEP StopPump_CIP4_01:
    _aStopPump_CIP4_01_entry(P1);  // entry action
END_STEP
TRANSITION FROM StopPump_CIP4_01 TO Tank_LowLevel_CIP4_01
    := TRUE;
END_TRANSITION
TRANSITION FROM Sprinkler_Request_CIP4 TO Tank_LowLevel_CIP4_02
    := TRUE;
END_TRANSITION
STEP Tank_LowLevel_CIP4_02:
    _aTank_LowLevel_CIP4_02_entry(P1);  // entry action
    _aTank_LowLevel_CIP4_02_active(N);  // step action
END_STEP
TRANSITION FROM Tank_LowLevel_CIP4_02 TO CIP4_Conn_Sprinkler
    := bStepDone;
END_TRANSITION
STEP CIP4_Conn_Sprinkler:
    _aCIP4_Conn_Sprinkler_entry(P1);  // entry action
    _aCIP4_Conn_Sprinkler_active(N);  // step action
END_STEP
TRANSITION FROM CIP4_Conn_Sprinkler TO ReadyToCondition_Count
    := bStepDone;
END_TRANSITION
TRANSITION FROM Condition_CIP4_Client TO StopPump_CIP4_02
    := bCIP_Condition_Failed;
END_TRANSITION
STEP StopPump_CIP4_02:
    _aStopPump_CIP4_02_entry(P1);  // entry action
END_STEP
TRANSITION FROM StopPump_CIP4_02 TO ReFill_Water_T94
    := TRUE;
END_TRANSITION
STEP ReFill_Water_T94:
    _aReFill_Water_T94_active(N);  // step action
END_STEP
TRANSITION FROM ReFill_Water_T94 TO Condition_CIP4_Client
    := bStepDone;
END_TRANSITION
STEP Tank_LowLevel_CIP4_01:
    _aTank_LowLevel_CIP4_01_active(N);  // step action
END_STEP
TRANSITION FROM Tank_LowLevel_CIP4_01 TO CIP4_Done
    := bStepDone;
END_TRANSITION
STEP CIP4_Done:  // min time T#2s
    _aCIP4_Done_entry(P1);  // entry action
END_STEP
TRANSITION FROM CIP4_Done TO End_Check
    := TRUE;
END_TRANSITION
STEP End_Check:
    _aEnd_Check_active(N);  // step action
END_STEP
TRANSITION FROM End_Check TO Disconnect_n_Drain_CIP_Client
    := bStepDone;
END_TRANSITION
TRANSITION FROM End_Check TO Get_Client
    := TRUE;
END_TRANSITION
STEP Disconnect_n_Drain_CIP_Client:
    _aDisconnect_n_Drain_CIP_Client_entry(P1);  // entry action
    _aDisconnect_n_Drain_CIP_Client_active(N);  // step action
END_STEP
TRANSITION FROM Disconnect_n_Drain_CIP_Client TO Done
    := bStepDone;
END_TRANSITION
STEP Done:  // min time T#0.1s
    _aDone_entry(P1);  // entry action
END_STEP
TRANSITION FROM Done TO Disconnect_Old_Client
    := TRUE;
END_TRANSITION
// branch label Branch28_act_Oper
// branch label Branch29_act_Oper
// branch label Branch27_act_Oper
// branch label Branch26_act_Oper
// branch label Branch0_act_Oper
// branch label Branch11_act_Oper
// branch label Branch10_act_Oper
// branch label Branch15_act_Oper
// branch label Branch14_act_Oper
// branch label Branch10_act_Oper_2
// branch label Branch23_act_Oper
// branch label Branch12_act_Oper
// branch label Branch9_act_Oper
// branch label Branch17_act_Oper
// branch label Branch18_act_Oper
// branch label Branch19_act_Oper
// branch label Branch24_act_Oper
// branch label Branch20_act_Oper
// branch label Branch8_act_Oper
// branch label Branch2_act_Oper
// branch label Branch3_act_Oper
END_ACTION

ACTION act_ReqBuffer:
rtPosMoveHMI_Up(Q=>);
IF rtPosMoveHMI_Up.Q THEN;
	m_PosMove_Up_HMI();
END_IF
rtPosMoveHMI_Down(Q=>);
IF rtPosMoveHMI_Down.Q THEN;
	m_PosMove_Down_HMI();
END_IF
rtPosDeleteHMI(Q=>);
IF rtPosDeleteHMI.Q THEN;
	m_PosDelete_HMI();
END_IF
rtPosDeleteAllHMI(Q=>);
IF rtPosDeleteAllHMI.Q THEN;
	m_PosDeleteAll_HMI();
END_IF

rtReqLocalCIP_Full_HMI(Q=>);
IF rtReqLocalCIP_Full_HMI.Q THEN;
	eReqLocal.eClient:=E_CIP_Usage.eLocal;
	eReqLocal.eType:=E_CIP_Type.Full;
	m_TakePosInCIPBuffer(stCIP_Request:=eReqLocal);
END_IF

rtReqLocalCIP_Detergent_HMI(Q=>);
IF rtReqLocalCIP_Detergent_HMI.Q THEN;
	eReqLocal.eClient:=E_CIP_Usage.eLocal;
	eReqLocal.eType:=E_CIP_Type.Detergent;
	m_TakePosInCIPBuffer(stCIP_Request:=eReqLocal);
END_IF

rtReqCleanEmpty_HMI(Q=>);
IF rtReqCleanEmpty_HMI.Q THEN;
	m_CleanEmpty_Spaces();
END_IF
END_ACTION

ACTION act_Run:
IF __ISVALIDREF(eRefClient_fbElement) THEN
	IF eRefClient_fbElement.bError AND SFCCurrentStep<>'Ready' THEN;
		m_Set_LastStepBeforeError();
		sError_Message:='Client Error';
		//mResetCycle();
	END_IF	
END_IF
END_ACTION

ACTION act_SprinklerCondition:


IF __ISVALIDREF(eRefClient_fbElement) THEN;
	IF TRUE
	AND eRefClient_fbElement.eState_Long>=E_Element_State_Long.eCIP_1_Rinzed 
	AND eRefClient_fbElement.eState_Long<=E_Element_State_Long.eCIP_2_Deterged 
	THEN;
		IF NOT bSprinkler THEN // Pipe
			tConditionTime	:=st_CIP_Param.t_ConditionDetergent;
			fFlowRate		:=st_CIP_Param.r_Flow_Pipe;
		ELSE // Sprinkler
			tConditionTime	:=st_CIP_Param.t_ConditionDetergent_Sprinkler;
			fFlowRate		:=st_CIP_Param.r_Flow_Sprinkler;
		END_IF	
		//rVolume_Collect :=st_CIP_Param.r_Volume_Collect_Detergent;
		//rVolume_Drain	:=st_CIP_Param.r_Volume_Drain_Detergent;
		//rVolume_Recycle	:=st_CIP_Param.r_Volume_Recycle_Detergent;
		
	ELSIF TRUE
	AND eRefClient_fbElement.eState_Long>=E_Element_State_Long.eCIP_3_Deterged_Clean 
	AND eRefClient_fbElement.eState_Long<=E_Element_State_Long.eCIP_4_Sanitized 
	THEN;
		IF NOT bSprinkler THEN // Pipe
			tConditionTime	:=st_CIP_Param.t_ConditionDisInfection;
			fFlowRate		:=st_CIP_Param.r_Flow_Pipe;
		ELSE // Sprinkler
			tConditionTime	:=st_CIP_Param.t_ConditionDisInfection_Sprinkler;
			fFlowRate		:=st_CIP_Param.r_Flow_Sprinkler;
		END_IF	
		//rVolume_Collect :=st_CIP_Param.r_Volume_Collect_DisInfection;
		//rVolume_Drain	:=st_CIP_Param.r_Volume_Drain_DisInfection;
		//rVolume_Recycle	:=st_CIP_Param.r_Volume_Recycle_DisInfection;
	END_IF	
END_IF
END_ACTION

ACTION act_ValveUpLow_Cntrl:
tOn(IN:= , PT:=T#1S , Q=> , ET=> );
tOff(IN:= , PT:=T#3S , Q=> , ET=> );
nClient:=eCIP_Usage:=eReq.eClient;

//To be deleted just for testing
//***************************************************************************************
IF bClientTypeIs_Tank AND bSprinkler THEN;
	gCIP_ValvUL[1,1]:=E_Pis_Name.e0_not_in_use;
	gCIP_ValvUL[1,2]:=E_Pis_Name.V3017;
	gCIP_ValvUL[1,3]:=E_Pis_Name.V3023;
	gCIP_ValvUL[1,4]:=E_Pis_Name.e0_not_in_use;
	gCIP_ValvUL[1,5]:=E_Pis_Name.e0_not_in_use;
	gCIP_ValvUL[1,6]:=E_Pis_Name.e0_not_in_use;
																	
	gCIP_ValvUL[2,1]:=E_Pis_Name.e0_not_in_use;
	gCIP_ValvUL[2,2]:=E_Pis_Name.V3027;
	gCIP_ValvUL[2,3]:=E_Pis_Name.V3028;
	gCIP_ValvUL[2,4]:=E_Pis_Name.e0_not_in_use;
	gCIP_ValvUL[2,5]:=E_Pis_Name.e0_not_in_use;
	gCIP_ValvUL[2,6]:=E_Pis_Name.e0_not_in_use;
																	
	gCIP_ValvUL[3,1]:=E_Pis_Name.e0_not_in_use;
	gCIP_ValvUL[3,2]:=E_Pis_Name.e0_not_in_use;
	gCIP_ValvUL[3,3]:=E_Pis_Name.V4017;
	gCIP_ValvUL[3,4]:=E_Pis_Name.v4023;
	gCIP_ValvUL[3,5]:=E_Pis_Name.e0_not_in_use;
	gCIP_ValvUL[3,6]:=E_Pis_Name.e0_not_in_use;
																	
	gCIP_ValvUL[4,1]:=E_Pis_Name.e0_not_in_use;
	gCIP_ValvUL[4,2]:=E_Pis_Name.e0_not_in_use;
	gCIP_ValvUL[4,3]:=E_Pis_Name.V4027;
	gCIP_ValvUL[4,4]:=E_Pis_Name.V4028;
	gCIP_ValvUL[4,5]:=E_Pis_Name.e0_not_in_use;
	gCIP_ValvUL[4,6]:=E_Pis_Name.e0_not_in_use;	
ELSE;
	gCIP_ValvUL[1,1]:=E_Pis_Name.V3004;
	gCIP_ValvUL[1,2]:=E_Pis_Name.e0_not_in_use;
	gCIP_ValvUL[1,3]:=E_Pis_Name.e0_not_in_use;
	gCIP_ValvUL[1,4]:=E_Pis_Name.e0_not_in_use;
	gCIP_ValvUL[1,5]:=E_Pis_Name.e0_not_in_use;
	gCIP_ValvUL[1,6]:=E_Pis_Name.e0_not_in_use;
																	
	gCIP_ValvUL[2,1]:=E_Pis_Name.V3010;
	gCIP_ValvUL[2,2]:=E_Pis_Name.e0_not_in_use;
	gCIP_ValvUL[2,3]:=E_Pis_Name.e0_not_in_use;
	gCIP_ValvUL[2,4]:=E_Pis_Name.e0_not_in_use;
	gCIP_ValvUL[2,5]:=E_Pis_Name.e0_not_in_use;
	gCIP_ValvUL[2,6]:=E_Pis_Name.e0_not_in_use;
																	
	gCIP_ValvUL[3,1]:=E_Pis_Name.V4034;
	gCIP_ValvUL[3,2]:=E_Pis_Name.V4004;
	gCIP_ValvUL[3,3]:=E_Pis_Name.e0_not_in_use;
	gCIP_ValvUL[3,4]:=E_Pis_Name.e0_not_in_use;
	gCIP_ValvUL[3,5]:=E_Pis_Name.e0_not_in_use;
	gCIP_ValvUL[3,6]:=E_Pis_Name.e0_not_in_use;
																	
	gCIP_ValvUL[4,1]:=E_Pis_Name.V4033;
	gCIP_ValvUL[4,2]:=E_Pis_Name.V4010;
	gCIP_ValvUL[4,3]:=E_Pis_Name.e0_not_in_use;
	gCIP_ValvUL[4,4]:=E_Pis_Name.e0_not_in_use;
	gCIP_ValvUL[4,5]:=E_Pis_Name.e0_not_in_use;
	gCIP_ValvUL[4,6]:=E_Pis_Name.e0_not_in_use;	
END_IF
(*
	gCIP_ValvUL[1,1]:=E_Pis_Name.V3004;
	gCIP_ValvUL[1,2]:=E_Pis_Name.V3017;
	gCIP_ValvUL[1,3]:=E_Pis_Name.V3023;
	gCIP_ValvUL[1,4]:=E_Pis_Name.e0_not_in_use;
	gCIP_ValvUL[1,5]:=E_Pis_Name.e0_not_in_use;
	gCIP_ValvUL[1,6]:=E_Pis_Name.e0_not_in_use;
																	
	gCIP_ValvUL[2,1]:=E_Pis_Name.V3010;
	gCIP_ValvUL[2,2]:=E_Pis_Name.V3027;
	gCIP_ValvUL[2,3]:=E_Pis_Name.V3028;
	gCIP_ValvUL[2,4]:=E_Pis_Name.e0_not_in_use;
	gCIP_ValvUL[2,5]:=E_Pis_Name.e0_not_in_use;
	gCIP_ValvUL[2,6]:=E_Pis_Name.e0_not_in_use;
																	
	gCIP_ValvUL[3,1]:=E_Pis_Name.V4034;
	gCIP_ValvUL[3,2]:=E_Pis_Name.V4004;
	gCIP_ValvUL[3,3]:=E_Pis_Name.V4017;
	gCIP_ValvUL[3,4]:=E_Pis_Name.v4023;
	gCIP_ValvUL[3,5]:=E_Pis_Name.e0_not_in_use;
	gCIP_ValvUL[3,6]:=E_Pis_Name.e0_not_in_use;
																	
	gCIP_ValvUL[4,1]:=E_Pis_Name.V4033;
	gCIP_ValvUL[4,2]:=E_Pis_Name.V4010;
	gCIP_ValvUL[4,3]:=E_Pis_Name.V4027;
	gCIP_ValvUL[4,4]:=E_Pis_Name.V4028;
	gCIP_ValvUL[4,5]:=E_Pis_Name.e0_not_in_use;
	gCIP_ValvUL[4,6]:=E_Pis_Name.e0_not_in_use;
*)
																
gCIP_ValvUL[5,1]:=E_Pis_Name.V3113;
gCIP_ValvUL[5,2]:=E_Pis_Name.V3004;
gCIP_ValvUL[5,3]:=E_Pis_Name.V3010;
gCIP_ValvUL[5,4]:=E_Pis_Name.V3023;
gCIP_ValvUL[5,5]:=E_Pis_Name.V3028;
gCIP_ValvUL[5,6]:=E_Pis_Name.e0_not_in_use;
																
gCIP_ValvUL[6,1]:=E_Pis_Name.v2114;
gCIP_ValvUL[6,2]:=E_Pis_Name.V4004;
gCIP_ValvUL[6,3]:=E_Pis_Name.V4010;
gCIP_ValvUL[6,4]:=E_Pis_Name.V2116;
gCIP_ValvUL[6,5]:=E_Pis_Name.V4023;
gCIP_ValvUL[6,6]:=E_Pis_Name.V4028;
																
gCIP_ValvUL[7,1]:=E_Pis_Name.V3017;
gCIP_ValvUL[7,2]:=E_Pis_Name.V3027;
gCIP_ValvUL[7,3]:=E_Pis_Name.e0_not_in_use;
gCIP_ValvUL[7,4]:=E_Pis_Name.e0_not_in_use;
gCIP_ValvUL[7,5]:=E_Pis_Name.e0_not_in_use;
gCIP_ValvUL[7,6]:=E_Pis_Name.e0_not_in_use;

gCIP_ValvUL[8,1]:=E_Pis_Name.V4017;
gCIP_ValvUL[8,2]:=E_Pis_Name.v4027;
gCIP_ValvUL[8,3]:=E_Pis_Name.V2115;
gCIP_ValvUL[8,4]:=E_Pis_Name.V4034;
gCIP_ValvUL[8,5]:=E_Pis_Name.V4033;
gCIP_ValvUL[8,6]:=E_Pis_Name.e0_not_in_use;	

// set upper or lowwer
gCIP_ValvUL_Seat[1,1]:=0;
gCIP_ValvUL_Seat[1,2]:=1;
gCIP_ValvUL_Seat[1,3]:=1;
gCIP_ValvUL_Seat[1,4]:=0;
gCIP_ValvUL_Seat[1,5]:=0;
gCIP_ValvUL_Seat[1,6]:=0; // Client 1 eTank_1,

gCIP_ValvUL_Seat[2,1]:=0;
gCIP_ValvUL_Seat[2,2]:=1;
gCIP_ValvUL_Seat[2,3]:=1;
gCIP_ValvUL_Seat[2,4]:=0;
gCIP_ValvUL_Seat[2,5]:=0;
gCIP_ValvUL_Seat[2,6]:=0; // Client 2 eTank_2,
															
gCIP_ValvUL_Seat[3,1]:=0;
gCIP_ValvUL_Seat[3,2]:=0;
gCIP_ValvUL_Seat[3,3]:=1;
gCIP_ValvUL_Seat[3,4]:=1;
gCIP_ValvUL_Seat[3,5]:=0;
gCIP_ValvUL_Seat[3,6]:=0; // Client 3 eTank_3,
															
gCIP_ValvUL_Seat[4,1]:=0;
gCIP_ValvUL_Seat[4,2]:=0;
gCIP_ValvUL_Seat[4,3]:=1;
gCIP_ValvUL_Seat[4,4]:=1;
gCIP_ValvUL_Seat[4,5]:=0;
gCIP_ValvUL_Seat[4,6]:=0; // Client 4 eTank_4,
															
gCIP_ValvUL_Seat[5,1]:=0;
gCIP_ValvUL_Seat[5,2]:=1;
gCIP_ValvUL_Seat[5,3]:=1;
gCIP_ValvUL_Seat[5,4]:=0;
gCIP_ValvUL_Seat[5,5]:=0;
gCIP_ValvUL_Seat[5,6]:=0; // Client 5
															
gCIP_ValvUL_Seat[6,1]:=0;
gCIP_ValvUL_Seat[6,2]:=1;
gCIP_ValvUL_Seat[6,3]:=1;
gCIP_ValvUL_Seat[6,4]:=0;
gCIP_ValvUL_Seat[6,5]:=0;
gCIP_ValvUL_Seat[6,6]:=0; // Client 6
															
gCIP_ValvUL_Seat[7,1]:=0;
gCIP_ValvUL_Seat[7,2]:=0;
gCIP_ValvUL_Seat[7,3]:=0;
gCIP_ValvUL_Seat[7,4]:=0;
gCIP_ValvUL_Seat[7,5]:=0;
gCIP_ValvUL_Seat[7,6]:=0; // Client 7
									
gCIP_ValvUL_Seat[8,1]:=0;
gCIP_ValvUL_Seat[8,2]:=0;
gCIP_ValvUL_Seat[8,3]:=0;
gCIP_ValvUL_Seat[8,4]:=1;
gCIP_ValvUL_Seat[8,5]:=1;
gCIP_ValvUL_Seat[8,6]:=0; // Client 8 	
//***************************************************************************************											

CASE nStep_Vlv OF
	0:
		//waiting step
		IF bClean_MixProof 
		AND nClient<=8 
		AND nClient>0 
		AND (tonr_CIP_Condition.IN
			OR (bClientTypeIs_Tank AND bSprinkler))
		THEN
			bValveCleanDone:=FALSE;
			sState:='Busy';
			//nI_1_act_valve:=1;//active valve
			//nI_2_act_pulses:=1;//active number of pulses
			//nI_3_act_repeats:=1;//active number of retries
			tOn.IN:=FALSE;
			tOff.IN:=FALSE;
			nStep_Vlv:=1;
		ELSIF bClean_MixProof AND (nClient>8 OR nClient<=0) THEN
			nStep_Vlv:=999;
		END_IF
	1:
		bClean_MixProof:=FALSE;
		nI_2_act_pulses:=1; // 4 =>> 5 pulses
		
		IF nI_1_act_valve<=6 THEN;
			IF TRUE 
			AND gCIP_ValvUL[nClient,nI_1_act_valve]<E_Pis_Name.last 
			AND nI_1_act_valve<=nMaxValves THEN;
				IF gCIP_ValvUL[nClient,nI_1_act_valve]>E_Pis_Name.e0_not_in_use THEN;
					//existing step
					nStep_Vlv:=2;			
				ELSE;
					nI_1_act_valve:=nI_1_act_valve+1;
				END_IF
			ELSE
				//DONE
				nStep_Vlv:=10;
			END_IF		
		ELSE;
			nStep_Vlv:=10;	
		END_IF
		

		
	2:
		ActvValve:=gCIP_ValvUL[nClient,nI_1_act_valve];
		bSeatStatus:=gCIP_ValvUL_Seat[nClient,nI_1_act_valve];
		nStep_Vlv:=3;
	3:
		
		//Open Valve
			//
			
		IF bSeatStatus THEN
			//Upper
			g_Piston.stPis_U_L[ActvValve].req_Upper:=TRUE;
		ELSE
			//Lower 
			g_Piston.stPis_U_L[ActvValve].req_Lower:=TRUE;
		END_IF
			
		tOn.IN:=TRUE;
		tOff.IN:=FALSE;
		
		IF tOn.Q 
		AND ((g_Piston.stPis_U_L[ActvValve].st_Upper AND g_Piston.stPis_U_L[ActvValve].req_Upper)
				OR 
			(g_Piston.stPis_U_L[ActvValve].st_Lower AND g_Piston.stPis_U_L[ActvValve].req_Lower))
		THEN;
			nStep_Vlv:=4;
		END_IF
		
	4:
		//Close valve
			//
			
		IF bSeatStatus THEN
			//Upper
			g_Piston.stPis_U_L[ActvValve].req_Upper:=FALSE;
		ELSE
			//Lower 
			g_Piston.stPis_U_L[ActvValve].req_Lower:=FALSE;
		END_IF
			
		tOn.IN:=FALSE;
		tOff.IN:=TRUE;
		
		IF tOff.Q
		AND g_Piston.stPis_U_L[ActvValve].st_Released
		AND nI_2_act_pulses>=nNumOfPulses 
		THEN
			//fetch another valve
			IF nI_1_act_valve < nMaxValves THEN;
				nI_1_act_valve:=nI_1_act_valve+1;
				nStep_Vlv:=1;	
			ELSE;
				//DONE
				nStep_Vlv:=10;	
			END_IF

		ELSIF tOff.Q
		AND g_Piston.stPis_U_L[ActvValve].st_Released		
		AND nI_2_act_pulses<nNumOfPulses 
		AND TRUE THEN
			//return to open
			nI_2_act_pulses:=nI_2_act_pulses+1;
			nStep_Vlv:=3;
		END_IF
	10:
		IF nI_3_act_repeats<nNumOfRetries THEN
			//returnng to repeat
			nI_3_act_repeats:=nI_3_act_repeats+1;
			nI_1_act_valve:=1;
			nStep_Vlv:=1;
		ELSE
			//Done
			nStep_Vlv:=100;
		END_IF
	100:
		//Done
		bValveCleanDone:=TRUE;
		sState:='Done';
		nStep_Vlv:=0;
	999:
		//error incorrect Client number
		sState:='Error. Incorect Client name';
		
END_CASE 

IF nStep_Vlv<>0 
AND (NOT Ready.x)
AND (stOper[E_ModeZone.eCIP].iActOperation=E_OperationButtons.ePauseAll
	//OR (NOT tonr_CIP_Condition.IN AND NOT(bClientTypeIs_Tank AND bSprinkler)))
	OR ton_Concentration_Filter.ET>T#10S
	OR bCIP_Condition_Failed)
THEN;
	m_MixProof_Release_All();
	nStep_Vlv:=0;
END_IF
END_ACTION

METHOD m_Check_ProductionTank_Low_Level : BOOL
VAR_INPUT
END_VAR
IF TRUE
AND __ISVALIDREF(fbTank1.ref_fbTankSensors) 
AND __ISVALIDREF(fbTank2.ref_fbTankSensors) 
AND __ISVALIDREF(fbTank3.ref_fbTankSensors) 
AND __ISVALIDREF(fbTank4.ref_fbTankSensors) 
THEN;
	
	CASE eReq.eClient OF
		E_CIP_Usage.eTank_1:;
					IF NOT fbTank1.ref_fbTankSensors.senLL THEN;
						tonTankLowLevel.IN:=TRUE;
					ELSE;
						tonTankLowLevel.IN:=FALSE;
					END_IF
		E_CIP_Usage.eTank_2:;
					IF NOT fbTank2.ref_fbTankSensors.senLL THEN;
						tonTankLowLevel.IN:=TRUE;
					ELSE;
						tonTankLowLevel.IN:=FALSE;
					END_IF
		E_CIP_Usage.eTank_3:;
					IF NOT fbTank3.ref_fbTankSensors.senLL THEN;
						tonTankLowLevel.IN:=TRUE;
					ELSE;
						tonTankLowLevel.IN:=FALSE;
					END_IF
		E_CIP_Usage.eTank_4:;
					IF NOT fbTank4.ref_fbTankSensors.senLL THEN;
						tonTankLowLevel.IN:=TRUE;
					ELSE;
						tonTankLowLevel.IN:=FALSE;
					END_IF
		E_CIP_Usage.eLine_Marinada:;
		E_CIP_Usage.eLine_Color:;
		E_CIP_Usage.eTriBlender_Marinada,
		E_CIP_Usage.eTriBlender_Color:;
					
	END_CASE	
	
	tonTankLowLevel(PT:=T#2S);
	IF bClientTypeIs_Tank 
	AND tonTankLowLevel.Q
	THEN;
		m_Check_ProductionTank_Low_Level:=TRUE;
		fb_PumpClient.m_Stop();
	ELSIF NOT bClientTypeIs_Tank 
	THEN;
		m_Check_ProductionTank_Low_Level:=TRUE;
		fb_PumpClient.m_Stop();
	ELSE;
		m_Check_ProductionTank_Low_Level:=FALSE;
	END_IF
	
END_IF
END_METHOD

METHOD m_CleanEmpty_Spaces : BOOL
VAR_INPUT
END_VAR

VAR
	i: INT;
	j: INT;
	stCIP_Request_Empty: ST_CIP_Request;
END_VAR
FOR i:=0 TO 9 DO
	IF i<>0 OR NOT bRun THEN;
		IF arCIP_RequestBufer[i].eClient=E_CIP_Usage.eNotInUse THEN;
			FOR j:=i+1 TO 9 DO
				IF arCIP_RequestBufer[j].eClient<>E_CIP_Usage.eNotInUse THEN;
					arCIP_RequestBufer[i]:=arCIP_RequestBufer[j];
					arCIP_RequestBufer[j]:=stCIP_Request_Empty;
					EXIT;
				END_IF
			END_FOR
		END_IF		
	END_IF
END_FOR
END_METHOD

METHOD m_ClientTank_IsEmpty : BOOL
VAR_INPUT
END_VAR
IF __ISVALIDREF(ref_lvlTank_Client) 
AND bClientTypeIs_Tank
THEN;
	m_ClientTank_IsEmpty:=ref_lvlTank_Client.e_state=E_Tank_Level.eEmpty;
ELSE;
	m_ClientTank_IsEmpty:=TRUE;
END_IF
END_METHOD

METHOD m_ClientTank_Level_IsHigher_Then : BOOL
VAR_INPUT
	min_Level: REAL:=150.0;
END_VAR
IF __ISVALIDREF(ref_lvlTank_Client) 
AND bClientTypeIs_Tank
THEN;
	m_ClientTank_Level_IsHigher_Then:=ref_lvlTank_Client.rTankLevel>=min_Level;
ELSE;
	m_ClientTank_Level_IsHigher_Then:=FALSE;
END_IF
END_METHOD

METHOD m_DashState_activate : BOOL
VAR_INPUT
	stage		: E_CIP_DashStage_List;
END_VAR
	IF arCIP_DashStage_list[stage] = E_CIP_DashStage.eCIPStage_ToBeDone THEN;
		arCIP_DashStage_list[stage]:=E_CIP_DashStage.eCIPStage_Active;
		eCIP_DashStage_actual:=stage;
		sCIP_DashStage_actual:=TO_STRING(eCIP_DashStage_actual);	
		RETURN;
	END_IF

(*
FOR stage:=m_DashState_from() TO m_DashState_to() DO
	IF arCIP_DashStage_list[stage] = E_CIP_DashStage.eCIPStage_ToBeDone THEN;
		arCIP_DashStage_list[stage]:=E_CIP_DashStage.eCIPStage_Active;
		eCIP_DashStage_actual:=stage;
		sCIP_DashStage_actual:=TO_STRING(eCIP_DashStage_actual);	
		RETURN;
	END_IF
END_FOR
*)
END_METHOD

METHOD m_DashState_done : BOOL
VAR_INPUT
	stage	: E_CIP_DashStage_List;
END_VAR
IF arCIP_DashStage_list[stage] = E_CIP_DashStage.eCIPStage_Active THEN;
	arCIP_DashStage_list[stage]:=E_CIP_DashStage.eCIPStage_Done;
	RETURN;
END_IF

(*
FOR stage:=m_DashState_from() TO m_DashState_to() DO
	IF arCIP_DashStage_list[stage] = E_CIP_DashStage.eCIPStage_Active THEN;
		arCIP_DashStage_list[stage]:=E_CIP_DashStage.eCIPStage_Done;
		RETURN;
	END_IF
END_FOR
*)
END_METHOD

METHOD m_DashState_from : E_CIP_DashStage_List
VAR
	eActCIP_State	: E_Element_State_Long;
END_VAR
eActCIP_State:=eRefClient_fbElement.eState_Long;

CASE eActCIP_State OF
	E_Element_State_Long.eNotClean:;
		m_DashState_from:=E_CIP_DashStage_List.e01_CIP1_Client_Drain_Product_Rest_Pipe;	
		
	E_Element_State_Long.eCIP_1_Rinzed:;
		m_DashState_from:=E_CIP_DashStage_List.e03_CIP2_Local_Detergent_Fill;	
	
	E_Element_State_Long.eCIP_2_Deterged:;
		m_DashState_from:=E_CIP_DashStage_List.e08_CIP3_Detergent_Collect;	
	
	E_Element_State_Long.eCIP_3_Deterged_Clean:;
		m_DashState_from:=E_CIP_DashStage_List.e12_CIP4_Local_DisInfection_Fill;	
	
	E_Element_State_Long.eCIP_4_Sanitized:;
		m_DashState_from:=E_CIP_DashStage_List.e17_CIP5_DisInfection_Collect;	
	
ELSE;
	//???
		m_DashState_from:=E_CIP_DashStage_List.eLast;
END_CASE
END_METHOD

METHOD m_DashState_Get_ToBeDone_List : BOOL
VAR
	//eActCIP_State	: E_Element_State_Long;
	//eCIP_req		: ST_CIP_Request;	
	stage			: E_CIP_DashStage_List;
END_VAR
//eActCIP_State:=eRefClient_fbElement.eState_Long;
//eCIP_req:=eReq;

//init
FOR stage:=E_CIP_DashStage_List.e00_NotSelected TO E_CIP_DashStage_List.eLast DO
	arCIP_DashStage_list[stage]:=E_CIP_DashStage.eCIPStage_NotAvalable;
END_FOR

//Start done condition stages
FOR stage:=E_CIP_DashStage_List.e00_NotSelected TO m_DashState_from()-1 DO
	IF m_DashState_Sprinkler(stage:=stage) THEN;
		IF bClientTypeIs_Tank THEN;
			arCIP_DashStage_list[stage]:=E_CIP_DashStage.eCIPStage_Done;
		ELSE;
			arCIP_DashStage_list[stage]:=E_CIP_DashStage.eCIPStage_NotAvalable;
		END_IF
	ELSE;
		arCIP_DashStage_list[stage]:=E_CIP_DashStage.eCIPStage_Done;
	END_IF
END_FOR

// Request conditions
FOR stage:=m_DashState_from() TO m_DashState_to() DO
	IF m_DashState_Sprinkler(stage:=stage) THEN;
		IF bClientTypeIs_Tank THEN;
			arCIP_DashStage_list[stage]:=E_CIP_DashStage.eCIPStage_ToBeDone;
		ELSE;
			arCIP_DashStage_list[stage]:=E_CIP_DashStage.eCIPStage_NotAvalable;
		END_IF
	ELSE;
		arCIP_DashStage_list[stage]:=E_CIP_DashStage.eCIPStage_ToBeDone;
	END_IF
END_FOR

//Do not requested 
FOR stage:=m_DashState_to()+1 TO E_CIP_DashStage_List.eLast DO
	IF m_DashState_Sprinkler(stage:=stage) THEN;
		IF bClientTypeIs_Tank THEN;
			arCIP_DashStage_list[stage]:=E_CIP_DashStage.eCIPStage_NotInUse;
		ELSE;
			arCIP_DashStage_list[stage]:=E_CIP_DashStage.eCIPStage_NotAvalable;
		END_IF
	ELSE;
		arCIP_DashStage_list[stage]:=E_CIP_DashStage.eCIPStage_NotInUse;
	END_IF
END_FOR
END_METHOD

METHOD m_DashState_MixProof_set : BOOL
VAR_INPUT
END_VAR
IF NOT __ISVALIDREF(eRefClient_fbElement) THEN;
	RETURN;
END_IF
CASE eCIP_Usage OF
	E_CIP_Usage.eNotInUse,
	E_CIP_Usage.eLocal:;
		FOR i:=1 TO 6 DO
			g_HMI.arCIP_DashStage_MixProof[i].sName:='';
			g_HMI.arCIP_DashStage_MixProof[i].bUpper:=FALSE;
			g_HMI.arCIP_DashStage_MixProof[i].bLower:=FALSE;
			g_HMI.arCIP_DashStage_MixProof[i].bRunning:=FALSE;
			g_HMI.arCIP_DashStage_MixProof[i].bDone:=FALSE;
		END_FOR	
ELSE;
		FOR i:=1 TO 6 DO
			g_HMI.arCIP_DashStage_MixProof[i].sName:=TO_STRING(gCIP_ValvUL[eCIP_Usage,i]);
			g_HMI.arCIP_DashStage_MixProof[i].bUpper:=gCIP_ValvUL_Seat[eCIP_Usage,i];
			g_HMI.arCIP_DashStage_MixProof[i].bLower:=NOT gCIP_ValvUL_Seat[eCIP_Usage,i];
			g_HMI.arCIP_DashStage_MixProof[i].bRunning:= nI_1_act_valve=i AND nStep_Vlv<>0;
			g_HMI.arCIP_DashStage_MixProof[i].bDone:= (nI_1_act_valve>i AND TRUE) OR bValveCleanDone;
		END_FOR	
END_CASE
END_METHOD

METHOD m_DashState_Sprinkler : BOOL
VAR_INPUT
	stage: E_CIP_DashStage_List;
END_VAR
CASE stage OF 
	E_CIP_DashStage_List.e02_CIP1_Client_Drain_Product_Rest_Sprinkler,
	E_CIP_DashStage_List.e07_CIP2_Client_Detergent_Condition_Sprinkler,
	E_CIP_DashStage_List.e11_CIP3_Detergent_Clean_Sprinkler,
	E_CIP_DashStage_List.e16_CIP4_Client_DisInfection_Condition_Sprinkler,
	E_CIP_DashStage_List.e20_CIP5_DisInfection_Clean_Sprinkler:;
		m_DashState_Sprinkler:=TRUE;
ELSE;
		m_DashState_Sprinkler:=FALSE;
END_CASE
END_METHOD

METHOD m_DashState_to : E_CIP_DashStage_List
VAR
	eCIP_req		: ST_CIP_Request;
END_VAR
eCIP_req:=eReq;

CASE eCIP_req.eType OF
	E_CIP_Type.R_Water:;
		m_DashState_to:=E_CIP_DashStage_List.e02_CIP1_Client_Drain_Product_Rest_Sprinkler;
		
	E_CIP_Type.Detergent:;
		m_DashState_to:=E_CIP_DashStage_List.e11_CIP3_Detergent_Clean_Sprinkler;
	
	E_CIP_Type.Full:;
		m_DashState_to:=E_CIP_DashStage_List.e20_CIP5_DisInfection_Clean_Sprinkler;

ELSE;
	//???
		m_DashState_to:=E_CIP_DashStage_List.eLast;	
END_CASE
END_METHOD

METHOD m_DashState_ToString_convertion : BOOL
VAR_INPUT
END_VAR

VAR
	eDashboard_CIP_State: E_CIP_DashStage_List:=E_CIP_DashStage_List.eLast;
END_VAR
FOR eDashboard_CIP_State:=0 TO E_CIP_DashStage_List.eLast DO
	//g_HMI.arCIP_DashStage_list[eDashboard_CIP_State]:=E_CIP_DashStage.eCIPStage_NotInUse;
	g_HMI.arCIP_DashStage_string[eDashboard_CIP_State]:=TO_STRING(eDashboard_CIP_State);
END_FOR
END_METHOD

METHOD m_Disconnect_All_Client : BOOL
VAR
	i: E_Element_List;
END_VAR
FOR i:=E_Element_List.eTank_1 TO E_Element_List.eLine_Color DO
	IF g_Data.fbElement[i].m_Get_InterConnection()=E_InterConnection.ConnToCIP THEN;
		g_Data.fbElement[i].m_Disconnect();
	END_IF
END_FOR
END_METHOD

METHOD m_MeasureTimeToHMI : TIME
VAR_INPUT
END_VAR
IF SFCCurrentStep='measureDelay_CIP2_1' THEN;
	m_MeasureTimeToHMI:=measureDelay_CIP2_1.t;
	
ELSIF SFCCurrentStep='measureDelay_CIP2_2' THEN;
	m_MeasureTimeToHMI:=measureDelay_CIP2_2.t;
	
ELSIF SFCCurrentStep='measureDelay_CIP3_1' THEN;
	m_MeasureTimeToHMI:=measureDelay_CIP3_1.t;
	
ELSIF SFCCurrentStep='measureDelay_CIP3_2' THEN;
	m_MeasureTimeToHMI:=measureDelay_CIP3_2.t;

ELSE;
	m_MeasureTimeToHMI:=T#0S;
END_IF
END_METHOD

METHOD m_MixProof_Release_All : BOOL
VAR_INPUT
END_VAR
VAR
	i: INT;
	j: INT;
END_VAR
FOR i:=1 TO 8 DO
	FOR j:=1 TO 6 DO
		ActvValve:=gCIP_ValvUL[i,j];
		g_Piston.stPis_U_L[ActvValve].req_Lower:=FALSE;
		g_Piston.stPis_U_L[ActvValve].req_Upper:=FALSE;
	END_FOR
END_FOR


FOR i:=1 TO 8 DO
	FOR j:=1 TO 6 DO
		ActvValve:=gCIP_ValvUL[i,j];
		IF g_Piston.stPis_U_L[ActvValve].exist
		AND NOT g_Piston.stPis_U_L[ActvValve].st_Released THEN;
			m_MixProof_Release_All:=FALSE;
			RETURN;
		END_IF
	END_FOR
END_FOR

m_MixProof_Release_All:=TRUE;
END_METHOD

METHOD m_MixProof_run : BOOL
VAR_INPUT
END_VAR
IF bValveCleanDone THEN;
	m_MixProof_run:=TRUE;
	bClean_MixProof:=FALSE;
ELSE;
	bClean_MixProof:=TRUE;
END_IF

m_DashState_MixProof_set();
END_METHOD

METHOD m_MixProof_set : BOOL
VAR_INPUT
END_VAR
nI_1_act_valve:=1;//active valve
nI_2_act_pulses:=1;//active number of pulses
nI_3_act_repeats:=1;//active number of retries

bClean_MixProof:=FALSE;
bValveCleanDone:=FALSE;
END_METHOD

METHOD m_OverFlowCorrect : REAL
VAR_INPUT
	rTc		:	REAL	;//Target concentration
	rAv		:	REAL	;//Actual volume
	rAc		:	REAL	;//Actual concentration
END_VAR
//Calculating the additional valume of fresh water to dalute the concentration
IF rTc=0 THEN;
	m_OverFlowCorrect:=0;
ELSE;
	m_OverFlowCorrect:=((rAv*rAc/100)/(rTc/100))-(rAv*rAc/100)-rAv+(rAv*rAc/100);
END_IF
END_METHOD

METHOD m_PosDelete_HMI : BOOL
VAR_INPUT
END_VAR
VAR
	stCIP_Request_Empty: ST_CIP_Request;
END_VAR
IF iPosSelect_HMI>=0 AND iPosSelect_HMI<9 THEN;
	IF iPosSelect_HMI<>0 OR NOT bRun THEN;
		arCIP_RequestBufer[iPosSelect_HMI]:=stCIP_Request_Empty;
	END_IF		
END_IF
END_METHOD

METHOD m_PosDeleteAll_HMI : BOOL
VAR_INPUT
END_VAR
VAR
	stCIP_Request_Empty: ST_CIP_Request;
	i: INT;
END_VAR

FOR i:=0 TO 9 DO
	IF i<>0 OR NOT bRun THEN;
		arCIP_RequestBufer[i]:=stCIP_Request_Empty;
	END_IF	
END_FOR
END_METHOD

METHOD m_PosMove_Down_HMI : BOOL
VAR_INPUT
END_VAR
VAR
	stCIP_Request_Temp: ST_CIP_Request;
	i: INT;
END_VAR
IF iPosSelect_HMI>=0 AND iPosSelect_HMI<9 THEN;
	IF iPosSelect_HMI<>0 OR NOT bRun THEN;		
			IF ((arCIP_RequestBufer[iPosSelect_HMI].eType=E_CIP_Type.R_Water 
				AND (arCIP_RequestBufer[iPosSelect_HMI+1].eType=E_CIP_Type.Detergent 
				OR arCIP_RequestBufer[iPosSelect_HMI+1].eType=E_CIP_Type.Full)) 
			OR (arCIP_RequestBufer[iPosSelect_HMI].eType=E_CIP_Type.Detergent 				
				AND arCIP_RequestBufer[iPosSelect_HMI+1].eType=E_CIP_Type.Full))
			AND (arCIP_RequestBufer[iPosSelect_HMI+1].eClient=arCIP_RequestBufer[iPosSelect_HMI].eClient) 
			THEN
				;
			ELSE
				stCIP_Request_Temp:=arCIP_RequestBufer[iPosSelect_HMI+1];
				arCIP_RequestBufer[iPosSelect_HMI+1]:=arCIP_RequestBufer[iPosSelect_HMI];
				arCIP_RequestBufer[iPosSelect_HMI]:=stCIP_Request_Temp;
				iPosSelect_HMI:=iPosSelect_HMI+1;	
			END_IF	
	END_IF
END_IF
END_METHOD

METHOD m_PosMove_Up_HMI : BOOL
VAR_INPUT
END_VAR
VAR
	stCIP_Request_Temp: ST_CIP_Request;
	i: INT;
	m: bool;
END_VAR
IF iPosSelect_HMI>0 AND iPosSelect_HMI<=9 THEN;
	IF iPosSelect_HMI<>1 OR NOT bRun THEN;			
			IF ((arCIP_RequestBufer[iPosSelect_HMI].eType=e_cip_type.Full 
				AND (arCIP_RequestBufer[iPosSelect_HMI-1].eType=E_CIP_Type.Detergent 
				OR arCIP_RequestBufer[iPosSelect_HMI-1].eType=E_CIP_Type.R_Water)) 
			OR (arCIP_RequestBufer[iPosSelect_HMI].eType=E_CIP_Type.Detergent 
				AND arCIP_RequestBufer[iPosSelect_HMI-1].eType=E_CIP_Type.R_Water))
			AND (arCIP_RequestBufer[iPosSelect_HMI-1].eClient=arCIP_RequestBufer[iPosSelect_HMI].eClient) 
			THEN
				;
			ELSE
				stCIP_Request_Temp:=arCIP_RequestBufer[iPosSelect_HMI-1];
				arCIP_RequestBufer[iPosSelect_HMI-1]:=arCIP_RequestBufer[iPosSelect_HMI];
				arCIP_RequestBufer[iPosSelect_HMI]:=stCIP_Request_Temp;
				iPosSelect_HMI:=iPosSelect_HMI-1;
			END_IF	
	END_IF
END_IF
END_METHOD

METHOD m_Set_SFCFlags_Reference : BOOL
//Set reference to SFC flags

refSFC.SFCInit REF= SFCInit;
refSFC.SFCReset REF= SFCReset;
refSFC.SFCError REF= SFCError;
refSFC.SFCEnableLimit REF= SFCEnableLimit;
refSFC.SFCErrorStep REF= SFCErrorStep;
refSFC.SFCErrorPOU REF= SFCErrorPOU;
refSFC.SFCQuitError REF= SFCQuitError;
refSFC.SFCPause REF= SFCPause;
refSFC.SFCTrans REF= SFCTrans;
refSFC.SFCCurrentStep REF= SFCCurrentStep;
refSFC.SFCTip REF= SFCTip;
refSFC.SFCTipMode REF= SFCTipMode;

// Cycle handle for SFC
m_SFC_Handle();

m_Set_Mode_Reference(inMoedeZone:=E_ModeZone.eCIP);
END_METHOD

METHOD m_Stirrer_production_tank : BOOL
VAR_INPUT
END_VAR


IF TRUE
//AND fbCIP_Source.m_CheckStatus(eReqStatus:=E_CIP_Source.eT93_R_Water) 
AND fbCIP_Usage.m_CheckStatus(eReqStatus:=eReq.eClient)
AND mCIP_Clients_status(command:=E_CIP_Client_Command.eCIP)
THEN
	fbTank1.cip_Pump_linked:=fbCIP_ClientTank_Marinade.m_CheckStatus(eReqStatus:=E_CIP_ClientTank.eTank_A);
	fbTank2.cip_Pump_linked:=fbCIP_ClientTank_Marinade.m_CheckStatus(eReqStatus:=E_CIP_ClientTank.eTank_B);
	fbTank3.cip_Pump_linked:=fbCIP_ClientTank_Color.m_CheckStatus(eReqStatus:=E_CIP_ClientTank.eTank_A);
	fbTank4.cip_Pump_linked:=fbCIP_ClientTank_Color.m_CheckStatus(eReqStatus:=E_CIP_ClientTank.eTank_B);

	CASE eReq.eClient OF	
		E_CIP_Usage.eTank_1:;
		E_CIP_Usage.eTank_2:;
		E_CIP_Usage.eTank_3:;					
		E_CIP_Usage.eTank_4:;
	ELSE;				
	END_CASE
ELSE;
	fbTank1.cip_Pump_linked:=FALSE;
	fbTank2.cip_Pump_linked:=FALSE;
	fbTank3.cip_Pump_linked:=FALSE;
	fbTank4.cip_Pump_linked:=FALSE;	
END_IF
END_METHOD

METHOD m_TakePosInCIPBuffer : BOOL
VAR_INPUT
	stCIP_Request: ST_CIP_Request;
END_VAR

VAR
	i: INT;
	m: bool;	
END_VAR
IF stCIP_Request.eClient<>E_CIP_Usage.eNotInUse
AND stCIP_Request.eType<>E_CIP_Type.NotSelected
AND g_data.fbElement[stCIP_Request.eClient].ProdStatus<>E_Prod_Status.Active
AND g_data.fbElement[stCIP_Request.eClient].eState_Long>E_Element_State_Long.eStandby 
AND ((stCIP_Request.eType=E_CIP_Type.R_Water AND g_data.fbElement[stCIP_Request.eClient].eState_Long<E_Element_State_Long.eCIP_1_Rinzed)
	OR (stCIP_Request.eType=E_CIP_Type.Detergent AND g_data.fbElement[stCIP_Request.eClient].eState_Long<E_Element_State_Long.eCIP_3_Deterged_Clean)
	OR (stCIP_Request.eType=E_CIP_Type.Full AND g_data.fbElement[stCIP_Request.eClient].eState_Long<E_Element_State_Long.eCIP_5_Done))

THEN
	FOR i:=0 TO 9 DO
		IF arCIP_RequestBufer[i].eClient=stCIP_Request.eClient 
			AND arCIP_RequestBufer[i].eType>=stCIP_Request.eType 
		THEN 	
				m:=FALSE;
				EXIT;
			ELSE
				m:=TRUE;
		END_IF
	END_FOR	
	IF m=TRUE THEN
		FOR i:=0 TO 9 DO
			IF arCIP_RequestBufer[i].eClient=E_CIP_Usage.eNotInUse 
			THEN;
				arCIP_RequestBufer[i]:=stCIP_Request;
				m:=FALSE;
				EXIT;
			END_IF
		END_FOR	
	END_IF
ELSIF stCIP_Request.eClient=E_CIP_Usage.eLocal
AND stCIP_Request.eType<>E_CIP_Type.NotSelected
THEN;
		FOR i:=0 TO 9 DO
			IF arCIP_RequestBufer[i].eClient=E_CIP_Usage.eNotInUse 
			THEN;
				arCIP_RequestBufer[i]:=stCIP_Request;
				m:=FALSE;
				EXIT;
			END_IF
		END_FOR		
END_IF
END_METHOD

METHOD mCIP_Clients_command : BOOL
VAR_INPUT
	command: E_CIP_Client_Command ;
END_VAR

//eReq.eClient<>E_CIP_Usage.eLocal
IF command=E_CIP_Client_Command.eDrain THEN;
	CASE eReq.eClient OF
		E_CIP_Usage.eTank_1:;
			g_Data.fbTankTarget_1.m_Run(eReqProc:=E_Tank_Target.eDrain);
		E_CIP_Usage.eTank_2:;
			g_Data.fbTankTarget_2.m_Run(eReqProc:=E_Tank_Target.eDrain);	
		E_CIP_Usage.eTank_3:;
			g_Data.fbTankTarget_3.m_Run(eReqProc:=E_Tank_Target.eDrain);	
		E_CIP_Usage.eTank_4:;
			g_Data.fbTankTarget_4.m_Run(eReqProc:=E_Tank_Target.eDrain);	
		E_CIP_Usage.eTriBlender_Marinada:;
			g_Data.fbTriBlenderSource_Marinade.m_Run(eReqProc:=E_Line_Source.eDrain);	
			g_Data.fbTriBlenderTarget_Marinade.m_Run(eReqProc:=E_Line_Target.eDrain);	
		E_CIP_Usage.eTriBlender_Color:;
			g_Data.fbTriBlenderSource_Color.m_Run(eReqProc:=E_Line_Source.eDrain);	
			g_Data.fbTriBlenderTarget_Color.m_Run(eReqProc:=E_Line_Target.eDrain);		
		E_CIP_Usage.eLine_Marinada:;
			g_Data.fbLineSource_Marinade.m_Run(eReqProc:=E_Line_Source.eDrain);	
			g_Data.fbLineTarget_Marinade.m_Run(eReqProc:=E_Line_Target.eDrain);	
		E_CIP_Usage.eLine_Color:;
			g_Data.fbLineSource_Color.m_Run(eReqProc:=E_Line_Source.eDrain);	
			g_Data.fbLineTarget_Color.m_Run(eReqProc:=E_Line_Target.eDrain);	
	ELSE;
		//wrong, - local
	END_CASE	
ELSIF command=E_CIP_Client_Command.eCIP THEN;
	CASE eReq.eClient OF
		E_CIP_Usage.eTank_1:;
			g_Data.fbTankTarget_1.m_Run(eReqProc:=E_Tank_Target.eCIP);
		E_CIP_Usage.eTank_2:;
			g_Data.fbTankTarget_2.m_Run(eReqProc:=E_Tank_Target.eCIP);	
		E_CIP_Usage.eTank_3:;
			g_Data.fbTankTarget_3.m_Run(eReqProc:=E_Tank_Target.eCIP);	
		E_CIP_Usage.eTank_4:;
			g_Data.fbTankTarget_4.m_Run(eReqProc:=E_Tank_Target.eCIP);	
		E_CIP_Usage.eTriBlender_Marinada:;
			g_Data.fbTriBlenderSource_Marinade.m_Run(eReqProc:=E_Line_Source.eCIP);	
			g_Data.fbTriBlenderTarget_Marinade.m_Run(eReqProc:=E_Line_Target.eCIP);	
		E_CIP_Usage.eTriBlender_Color:;
			g_Data.fbTriBlenderSource_Color.m_Run(eReqProc:=E_Line_Source.eCIP);	
			g_Data.fbTriBlenderTarget_Color.m_Run(eReqProc:=E_Line_Target.eCIP);		
		E_CIP_Usage.eLine_Marinada:;
			g_Data.fbLineSource_Marinade.m_Run(eReqProc:=E_Line_Source.eCIP);	
			g_Data.fbLineTarget_Marinade.m_Run(eReqProc:=E_Line_Target.eCIP);	
		E_CIP_Usage.eLine_Color:;
			g_Data.fbLineSource_Color.m_Run(eReqProc:=E_Line_Source.eCIP);	
			g_Data.fbLineTarget_Color.m_Run(eReqProc:=E_Line_Target.eCIP);	
	ELSE;
		//wrong, - local
	END_CASE	
END_IF
END_METHOD

METHOD mCIP_Clients_status : BOOL
VAR_INPUT
	command: E_CIP_Client_Command ;
END_VAR

//eReq.eClient<>E_CIP_Usage.eLocal
IF command=E_CIP_Client_Command.eDrain THEN;
	CASE eReq.eClient OF
		E_CIP_Usage.eTank_1:;
			IF g_Data.fbTankTarget_1.m_CheckStatus(eReqStatus:=E_Tank_Target.eDrain) THEN;
				mCIP_Clients_status:=TRUE;
			ELSE;
				mCIP_Clients_status:=FALSE;	
			END_IF
		E_CIP_Usage.eTank_2:;
			IF g_Data.fbTankTarget_2.m_CheckStatus(eReqStatus:=E_Tank_Target.eDrain) THEN;
				mCIP_Clients_status:=TRUE;
			ELSE;
				mCIP_Clients_status:=FALSE;	
			END_IF	
		E_CIP_Usage.eTank_3:;
			IF g_Data.fbTankTarget_3.m_CheckStatus(eReqStatus:=E_Tank_Target.eDrain) THEN;
				mCIP_Clients_status:=TRUE;
			ELSE;
				mCIP_Clients_status:=FALSE;	
			END_IF	
		E_CIP_Usage.eTank_4:;
			IF g_Data.fbTankTarget_4.m_CheckStatus(eReqStatus:=E_Tank_Target.eDrain) THEN;
				mCIP_Clients_status:=TRUE;
			ELSE;
				mCIP_Clients_status:=FALSE;	
			END_IF	
		E_CIP_Usage.eTriBlender_Marinada:;
			IF  g_Data.fbTriBlenderSource_Marinade.m_CheckStatus(eReqStatus:=E_Line_Source.eDrain) 
			AND g_Data.fbTriBlenderTarget_Marinade.m_CheckStatus(eReqStatus:=E_Line_Target.eDrain) THEN;
				mCIP_Clients_status:=TRUE;
			ELSE;
				mCIP_Clients_status:=FALSE;	
			END_IF
		E_CIP_Usage.eTriBlender_Color:;
			IF  g_Data.fbTriBlenderSource_Color.m_CheckStatus(eReqStatus:=E_Line_Source.eDrain) 
			AND g_Data.fbTriBlenderTarget_Color.m_CheckStatus(eReqStatus:=E_Line_Target.eDrain) THEN;
				mCIP_Clients_status:=TRUE;
			ELSE;
				mCIP_Clients_status:=FALSE;	
			END_IF		
		E_CIP_Usage.eLine_Marinada:;
			IF  g_Data.fbLineSource_Marinade.m_CheckStatus(eReqStatus:=E_Line_Source.eDrain) 
			AND g_Data.fbLineTarget_Marinade.m_CheckStatus(eReqStatus:=E_Line_Target.eDrain) THEN;
				mCIP_Clients_status:=TRUE;
			ELSE;
				mCIP_Clients_status:=FALSE;	
			END_IF	
		E_CIP_Usage.eLine_Color:;
			IF  g_Data.fbLineSource_Color.m_CheckStatus(eReqStatus:=E_Line_Source.eDrain) 
			AND g_Data.fbLineTarget_Color.m_CheckStatus(eReqStatus:=E_Line_Target.eDrain) THEN;
				mCIP_Clients_status:=TRUE;
			ELSE;
				mCIP_Clients_status:=FALSE;	
			END_IF	
	ELSE;// local
		mCIP_Clients_status:=TRUE;
	END_CASE	
ELSIF command=E_CIP_Client_Command.eCIP THEN;
	CASE eReq.eClient OF
		E_CIP_Usage.eTank_1:;
			IF g_Data.fbTankTarget_1.m_CheckStatus(eReqStatus:=E_Tank_Target.eCIP) THEN;
				mCIP_Clients_status:=TRUE;
			ELSE;
				mCIP_Clients_status:=FALSE;	
			END_IF
		E_CIP_Usage.eTank_2:;
			IF g_Data.fbTankTarget_2.m_CheckStatus(eReqStatus:=E_Tank_Target.eCIP) THEN;
				mCIP_Clients_status:=TRUE;
			ELSE;
				mCIP_Clients_status:=FALSE;	
			END_IF	
		E_CIP_Usage.eTank_3:;
			IF g_Data.fbTankTarget_3.m_CheckStatus(eReqStatus:=E_Tank_Target.eCIP) THEN;
				mCIP_Clients_status:=TRUE;
			ELSE;
				mCIP_Clients_status:=FALSE;	
			END_IF	
		E_CIP_Usage.eTank_4:;
			IF g_Data.fbTankTarget_4.m_CheckStatus(eReqStatus:=E_Tank_Target.eCIP) THEN;
				mCIP_Clients_status:=TRUE;
			ELSE;
				mCIP_Clients_status:=FALSE;	
			END_IF	
		E_CIP_Usage.eTriBlender_Marinada:;
			IF  g_Data.fbTriBlenderSource_Marinade.m_CheckStatus(eReqStatus:=E_Line_Source.eCIP) 
			AND g_Data.fbTriBlenderTarget_Marinade.m_CheckStatus(eReqStatus:=E_Line_Target.eCIP) THEN;
				mCIP_Clients_status:=TRUE;
			ELSE;
				mCIP_Clients_status:=FALSE;	
			END_IF
		E_CIP_Usage.eTriBlender_Color:;
			IF  g_Data.fbTriBlenderSource_Color.m_CheckStatus(eReqStatus:=E_Line_Source.eCIP) 
			AND g_Data.fbTriBlenderTarget_Color.m_CheckStatus(eReqStatus:=E_Line_Target.eCIP) THEN;
				mCIP_Clients_status:=TRUE;
			ELSE;
				mCIP_Clients_status:=FALSE;	
			END_IF		
		E_CIP_Usage.eLine_Marinada:;
			IF  g_Data.fbLineSource_Marinade.m_CheckStatus(eReqStatus:=E_Line_Source.eCIP) 
			AND g_Data.fbLineTarget_Marinade.m_CheckStatus(eReqStatus:=E_Line_Target.eCIP) THEN;
				mCIP_Clients_status:=TRUE;
			ELSE;
				mCIP_Clients_status:=FALSE;	
			END_IF	
		E_CIP_Usage.eLine_Color:;
			IF  g_Data.fbLineSource_Color.m_CheckStatus(eReqStatus:=E_Line_Source.eCIP) 
			AND g_Data.fbLineTarget_Color.m_CheckStatus(eReqStatus:=E_Line_Target.eCIP) THEN;
				mCIP_Clients_status:=TRUE;
			ELSE;
				mCIP_Clients_status:=FALSE;	
			END_IF	
	ELSE;// local
		mCIP_Clients_status:=TRUE;
	END_CASE	
	
ELSIF command=E_CIP_Client_Command.eClose THEN;
	CASE eReq.eClient OF
		E_CIP_Usage.eTank_1:;
			IF g_Data.fbTankTarget_1.m_CheckStatus(eReqStatus:=E_Tank_Target.eClose) THEN;
				mCIP_Clients_status:=TRUE;
			ELSE;
				mCIP_Clients_status:=FALSE;	
			END_IF
		E_CIP_Usage.eTank_2:;
			IF g_Data.fbTankTarget_2.m_CheckStatus(eReqStatus:=E_Tank_Target.eClose) THEN;
				mCIP_Clients_status:=TRUE;
			ELSE;
				mCIP_Clients_status:=FALSE;	
			END_IF	
		E_CIP_Usage.eTank_3:;
			IF g_Data.fbTankTarget_3.m_CheckStatus(eReqStatus:=E_Tank_Target.eClose) THEN;
				mCIP_Clients_status:=TRUE;
			ELSE;
				mCIP_Clients_status:=FALSE;	
			END_IF	
		E_CIP_Usage.eTank_4:;
			IF g_Data.fbTankTarget_4.m_CheckStatus(eReqStatus:=E_Tank_Target.eClose) THEN;
				mCIP_Clients_status:=TRUE;
			ELSE;
				mCIP_Clients_status:=FALSE;	
			END_IF	
		E_CIP_Usage.eTriBlender_Marinada:;
			IF  g_Data.fbTriBlenderSource_Marinade.m_CheckStatus(eReqStatus:=E_Line_Source.eClose) 
			AND g_Data.fbTriBlenderTarget_Marinade.m_CheckStatus(eReqStatus:=E_Line_Target.eClose) THEN;
				mCIP_Clients_status:=TRUE;
			ELSE;
				mCIP_Clients_status:=FALSE;	
			END_IF
		E_CIP_Usage.eTriBlender_Color:;
			IF  g_Data.fbTriBlenderSource_Color.m_CheckStatus(eReqStatus:=E_Line_Source.eClose) 
			AND g_Data.fbTriBlenderTarget_Color.m_CheckStatus(eReqStatus:=E_Line_Target.eClose) THEN;
				mCIP_Clients_status:=TRUE;
			ELSE;
				mCIP_Clients_status:=FALSE;	
			END_IF		
		E_CIP_Usage.eLine_Marinada:;
			IF  g_Data.fbLineSource_Marinade.m_CheckStatus(eReqStatus:=E_Line_Source.eClose) 
			AND g_Data.fbLineTarget_Marinade.m_CheckStatus(eReqStatus:=E_Line_Target.eClose) THEN;
				mCIP_Clients_status:=TRUE;
			ELSE;
				mCIP_Clients_status:=FALSE;	
			END_IF	
		E_CIP_Usage.eLine_Color:;
			IF  g_Data.fbLineSource_Color.m_CheckStatus(eReqStatus:=E_Line_Source.eClose) 
			AND g_Data.fbLineTarget_Color.m_CheckStatus(eReqStatus:=E_Line_Target.eClose) THEN;
				mCIP_Clients_status:=TRUE;
			ELSE;
				mCIP_Clients_status:=FALSE;	
			END_IF	
	ELSE;// local
		mCIP_Clients_status:=TRUE;
	END_CASE		
END_IF
END_METHOD

METHOD mFillWater : BOOL
VAR_INPUT
END_VAR

VAR
	reqVolume: REAL;	
	valve : E_Pis_Name;;
	actLevel: REAL;
	fillCondition: BOOL;	
	
END_VAR
IF TRUE 
AND fbPis.m_CheckByRecipe(stPis:=stPis_FillWater_T91, req:=E_Piston_Recipe_State.Release)
AND fbPis.m_CheckByRecipe(stPis:=stPis_FillWater_T92, req:=E_Piston_Recipe_State.Release)
AND fbPis.m_CheckByRecipe(stPis:=stPis_FillWater_T93, req:=E_Piston_Recipe_State.Release)
AND bStateSafe
AND MAIN.bTemp_Water_Overweight_check
THEN;
	fillCondition:=TRUE;
ELSE;
	fillCondition:=FALSE;
END_IF

reqVolume:=st_CIP_Param.r_Tank94_Volume;
IF g_Data.arr_CIP_Param[E_CIP_Usage.eLocal].r_Tank94_Volume>reqVolume THEN;
	reqVolume:=g_Data.arr_CIP_Param[E_CIP_Usage.eLocal].r_Tank94_Volume;
END_IF

fbHysteresisFillT94(
	fIn:= lvlTank_T94.rTankLevel, 
	fHigh:= reqVolume, 
	fLow:= reqVolume-50.0, 
	iDigitsAfterDot:= 1, 
	bOut=> );

IF eMode<>E_CIP_Mode.eOff THEN;
	IF fbPis.m_CheckByRecipe(stPis:=stPis_FillWater_T94, req:=E_Piston_Recipe_State.Act) 
	AND (NOT fbHysteresisFillT94.bOut
	OR NOT fillCondition)
	THEN;
		//stPis_FillWater_T94.req_Close:=TRUE;
		fbPis.m_SetByRecipe(stPis:=stPis_FillWater_T94, req:=E_Piston_Recipe_State.Release);
		
	ELSIF fbPis.m_CheckByRecipe(stPis:=stPis_FillWater_T94, req:=E_Piston_Recipe_State.Release) 
	AND fbHysteresisFillT94.bOut
	AND fillCondition
	THEN;
		IF NOT arrTanksSens[E_Tank_Name.T94].get_stTankLevel_OverFlow() THEN;
			fbPis.m_SetByRecipe(stPis:=stPis_FillWater_T94, req:=E_Piston_Recipe_State.Act);			
		END_IF	
	END_IF	
END_IF
	
	
(*
fbFillT94(	
		valve:= valFillWater_T94, 
		reqLevel:= reqVolume, 
		actLevel:= lvlTank_T94.rTankLevel, 
		fillCondition:= );
*)
END_METHOD

METHOD mLoadDefProcessSetPoints : BOOL
VAR_INPUT
END_VAR

	stDetergent.ToleranceHigh:=0.05;
	stDetergent.ToleravceLow:=0.05;
	stTemperature_Deterg.ToleranceHigh:=1;
	stTemperature_Deterg.ToleravceLow:=1;
	stDisInfectant.ToleranceHigh:=0.05;
	stDisInfectant.ToleravceLow:=0.05;
	stTemperature_Dis.ToleranceHigh:=1;//0.5
	stTemperature_Dis.ToleravceLow:=1;//0.5
	stFlow1_Rate.ToleranceHigh:=10;
	stFlow1_Rate.ToleravceLow:=10;
	stFlow2_Rate.ToleranceHigh:=10;
	stFlow2_Rate.ToleravceLow:=10;
	stColor_Level.ToleranceHigh:=10;
	stColor_Level.ToleravceLow:=10;
	stMarinada_Level.ToleranceHigh:=10;
	stMarinada_Level.ToleravceLow:=10;
	stP1001_Pressure.ToleranceHigh:=1;
	stP1001_Pressure.ToleravceLow:=1;
END_METHOD

METHOD mProcessDeviation : REAL
VAR_INPUT
	reqValue: REAL;
	processValue: REAL;
END_VAR
mProcessDeviation:=reqValue-processValue;
END_METHOD

METHOD mVolumeMeter : BOOL
VAR_INPUT
END_VAR
delta_T91_Volume:=lvlTank_T91.rTankLevel-memo_T91_Level_start;//de
delta_T92_Volume:=lvlTank_T92.rTankLevel-memo_T92_Level_start;
delta_T93_Volume:=lvlTank_T93.rTankLevel-memo_T93_Level_start;
delta_T94_Volume:=lvlTank_T94.rTankLevel-memo_T94_Level_start;
END_METHOD

METHOD mVolumeReset_All : BOOL
VAR_INPUT
END_VAR
memo_T91_Level_start:=lvlTank_T91.rTankLevel;
memo_T92_Level_start:=lvlTank_T92.rTankLevel;
memo_T93_Level_start:=lvlTank_T93.rTankLevel;
memo_T94_Level_start:=lvlTank_T94.rTankLevel;
END_METHOD

END_FUNCTION_BLOCK

// ---- 00 Library/13 Process Control/FB_ProcessControl.TcPOU
FUNCTION_BLOCK FB_ProcessControl

VAR_IN_OUT
	stProcessControl	:	ST_ProcessControl	;
END_VAR
VAR
	bRun			: BOOL	;
	//fbPID	: 	FB_BasicPID	;
	fbPID	: 	PID	;
	hystCIP_SetPoint: FB_Hysteresis_REAL;
	Call_ActDelayTON	: TON	;
	
	handling_PID_Manual: TON;

END_VAR

//stProcessControl.bManual:=TRUE;



Call_ActDelayTON(IN:=stProcessControl.bActiveCntr , PT:=T#1S , Q=> , ET=> );

m_Check();

act_Call_PID();
act_CallHyst();

handling_PID_Manual(PT:=T#0.5S);//, IN:=TRUE
IF handling_PID_Manual.Q THEN;
	stProcessControl.bManual:=TRUE;
ELSE;
	stProcessControl.bManual:=FALSE;
END_IF

ACTION act_Call_PID:
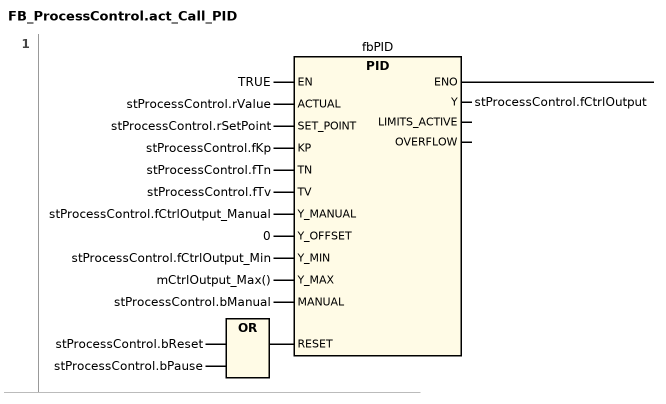
// NETWORK 1
fbPID(
    ACTUAL := stProcessControl.rValue,
    SET_POINT := stProcessControl.rSetPoint,
    KP := stProcessControl.fKp,
    TN := stProcessControl.fTn,
    TV := stProcessControl.fTv,
    Y_MANUAL := stProcessControl.fCtrlOutput_Manual,
    Y_OFFSET := 0,
    Y_MIN := stProcessControl.fCtrlOutput_Min,
    Y_MAX := mCtrlOutput_Max(),
    MANUAL := stProcessControl.bManual,
    RESET := stProcessControl.bReset OR stProcessControl.bPause,
    Y => stProcessControl.fCtrlOutput); // PID
END_ACTION

ACTION act_Call_PID_old:

	
(*
fbPID(
	fSetpointValue:=stProcessControl.rSetPoint , 
	fActualValue:=stProcessControl.rValue , 
	bReset:=stProcessControl.bReset , 
	fCtrlCycleTime:=stProcessControl.fCtrlCycleTime , 
	fKp:=stProcessControl.fKp , 
	fTn:=stProcessControl.fTn , 
	fTv:=stProcessControl.fTv , 
	fTd:=stProcessControl.fTd , 
	fCtrlOutput=>stProcessControl.fCtrlOutput , 
	nErrorStatus=>stProcessControl.nErrorStatus );
*)
END_ACTION

ACTION act_CallHyst:
hystCIP_SetPoint(
	fIn:=stProcessControl.rValue,//g_HMI.stT4_Sens.rTankLevel,
	fHigh:=stProcessControl.fHystHigh,
	fLow:=stProcessControl.fHystLow,
	iDigitsAfterDot:=,
	bOut=>stProcessControl.bHystOut);
END_ACTION

METHOD m_Check : BOOL
VAR_INPUT
END_VAR
IF bRun THEN 
	stProcessControl.bActiveCntr:=TRUE; 
ELSIF NOT bRun AND Call_ActDelayTON.Q THEN
	stProcessControl.bActiveCntr:=FALSE;
END_IF

IF bRun THEN
	stProcessControl.Deviation:=stProcessControl.rSetPoint-stProcessControl.rValue;
	stProcessControl.Control_ON:=FALSE;
	stProcessControl.OverFlow:=FALSE;
	stProcessControl.bDone:=FALSE;
	
	IF stProcessControl.Deviation >= stProcessControl.ToleravceLow THEN;
		//Value too low needs to be increased
		stProcessControl.Control_ON:=TRUE;
		stProcessControl.OverFlow:=FALSE;
		stProcessControl.bDone:=FALSE;
	ELSIF stProcessControl.Deviation <= -stProcessControl.ToleranceHigh THEN;
		//value too high need to be decreased
		stProcessControl.OverFlow:=TRUE;
		stProcessControl.Control_ON:=TRUE;
		stProcessControl.bDone:=FALSE;
		//message
	ELSE;
		// Done, value in tolerace
		stProcessControl.OverFlow:=FALSE;
		stProcessControl.Control_ON:=FALSE;
		stProcessControl.bDone:=TRUE;
	END_IF
	bRun:=FALSE;
END_IF
END_METHOD

METHOD mCtrlOutput_Max : REAL
VAR_INPUT
END_VAR

VAR
	span: LREAL;
END_VAR


span:=ABS(stProcessControl.fCtrlOutput_Max-stProcessControl.fCtrlOutput_Min);
//LimitedPrecentage:=
IF stProcessControl.rValue>stProcessControl.rValue_Min_To_ReleaseControl THEN;
	mCtrlOutput_Max:=stProcessControl.fCtrlOutput_Max;
ELSE;
	mCtrlOutput_Max:=stProcessControl.fCtrlOutput_Min+(span*0.3);
END_IF
END_METHOD

METHOD mPause : BOOL
VAR_INPUT
	value: BOOL;
END_VAR
stProcessControl.bPause:=value;
END_METHOD

METHOD mReset : BOOL
VAR_INPUT
END_VAR
stProcessControl.Control_ON:=FALSE;
stProcessControl.OverFlow:=FALSE;
stProcessControl.bDone:=FALSE;
END_METHOD

METHOD mRun : BOOL
VAR_INPUT
	//Set_Point: REAL;
END_VAR
bRun:=TRUE;
//stProcessControl.rSetPoint:=Set_Point;
m_Check();



mRun:=stProcessControl.bDone;
END_METHOD

METHOD mRun_Hyst : REAL
VAR_INPUT
END_VAR
stProcessControl.bManual:=FALSE;
IF stProcessControl.bHystOut THEN
	mRun_Hyst:=stProcessControl.rHystOutLow;
ELSE
	mRun_Hyst:=stProcessControl.rHystOutHigh;
END_IF
END_METHOD

METHOD mRun_PID : REAL
VAR_INPUT
	Set_Point: REAL;
	controlManual: BOOL;
END_VAR
mRun();//mRun(Set_Point:=Set_Point);
//stProcessControl.bManual:=controlManual;
//stProcessControl.rSetPoint:=Set_Point;
handling_PID_Manual(IN:=controlManual);
mRun_PID:=stProcessControl.fCtrlOutput;
END_METHOD

METHOD mRun_With_SP : BOOL
VAR_INPUT
	Set_Point: REAL;
END_VAR
stProcessControl.rSetPoint:=Set_Point;
bRun:=TRUE;
mRun();
stProcessControl.rSetPoint:=Set_Point;
mRun_With_SP:=stProcessControl.bDone;
END_METHOD

END_FUNCTION_BLOCK

// ---- 00 Library/10 Utils/FB_Hysteresis_REAL.TcPOU
FUNCTION_BLOCK FB_Hysteresis_REAL
VAR_INPUT
	fIn		: REAL; // in case of iDigitsAfterDot=2 max value 327.67 * 100 >> INTEGER Value limitation
	fHigh	: REAL;
	fLow	: REAL;
	iDigitsAfterDot: INT:=1; //min 0 , max 3

END_VAR
VAR_OUTPUT
	bOut	: BOOL;
END_VAR
VAR
	fbHys: HYSTERESIS;
	mult: INT;
	iDigitsAfterDot_Local: INT:=2; //min 0 , max 3


END_VAR

IF iDigitsAfterDot < 0 THEN;
	iDigitsAfterDot_Local:=0;
ELSIF iDigitsAfterDot > 3 THEN;
	iDigitsAfterDot_Local:=3;
ELSE;
	iDigitsAfterDot_Local:=iDigitsAfterDot;
END_IF
 

CASE iDigitsAfterDot_Local OF
	0:mult:=1;
	1:mult:=10;
	2:mult:=100;
	3:mult:=1000;
END_CASE

fbHys.HIGH:=REAL_TO_INT(fHigh*mult);
fbHys.LOW:=REAL_TO_INT(fLow*mult);
fbHys.IN:=REAL_TO_INT(fIn*mult);

fbHys(OUT=>bOut);

END_FUNCTION_BLOCK

// ---- 00 Library/10 Utils/TONR.TcPOU
FUNCTION_BLOCK TONR //Retentive Timer
VAR_INPUT
    IN : BOOL;         // Input signal
	ResetTime: BOOL;	//Reset Accumulating Time
    PT : TIME := T#0S; // Preset time
END_VAR
VAR_OUTPUT
    Q : BOOL;          // Output signal (true when time is reached)
    ET : TIME;         // Elapsed time
END_VAR
VAR
    StartTime : TIME := T#0S; // Start time storage
    IsTiming : BOOL := FALSE; // Timing state
END_VAR

// Start or continue timing when the input is true
IF IN THEN
    IF NOT IsTiming THEN
        StartTime := DT_TO_TIME(dtRealTime) - ET; // Adjust start time if resuming
        IsTiming := TRUE;
    END_IF
    ET := DT_TO_TIME(dtRealTime) - StartTime; // Calculate elapsed time
ELSE
    IsTiming := FALSE; // Stop timing but retain elapsed time
END_IF

IF ResetTime THEN
	ResetTime:=FALSE;
	IsTiming := FALSE; // Stop timing but retain elapsed time
	ET:=T#0s;
END_IF
 
// Check if the elapsed time has reached the preset time
IF ET >= PT THEN
    Q := TRUE;
ELSE
    Q := FALSE;
END_IF

END_FUNCTION_BLOCK

// ---- 03 Project/11 Tank/FB_ProductionTank.TcPOU
FUNCTION_BLOCK FB_ProductionTank EXTENDS FB_SFC_Cycle IMPLEMENTS ITF_FB_SFC_Cycle
VAR_INPUT
	eElementID		: E_Element_List;
	
	stTankValves				:	st_TankValves		;
	stLineSourceValves			:	st_LineSourceValves	;
	stTriBlenderSourceValves	:	st_LineSourceValves	;
	stLineTargetValves			:	st_LineTargetValves	;
	stfbTriBlenderTargetValves	:	st_LineTargetValves	;

	
	
	//valOutlet		: E_Pis_Name;//Comment?
	//valLine			: E_Pis_Name;//Comment?
	//valTriBlender	: E_Pis_Name;//Comment?
	//valDrain		: E_Pis_Name;//Comment?
	//valCIP			: E_Pis_Name;//Comment?
	
	valFilling				: E_Pis_Name;
	valFillWater			: E_Pis_Name;
	valFillWaterDrain		: E_Pis_Name;
	valDrainTapWater		: E_Pis_Name;
	
	eTank_Name				: E_Tank_Name;

	
	sens_TankTemp			: E_ASense_Name	;//Tenk temperature sensor ID
	
	valCW_In				:	E_Pis_Name	;//Valve to control tank temperature In
	valCW_Out				:	E_Pis_Name	;//Valve to control tank temperature Out (always at 100 open)
	
	//pumpEnum			:	E_Pump_List	;
	
END_VAR
VAR_OUTPUT
END_VAR
VAR
	sTank_Name			: STRING;
	refElement			: REFERENCE TO FB_Element;
	refState_Long		: REFERENCE TO E_Element_State_Long;
	eReq				: E_Request_List;		
	eProcess			: E_Element_Process;
	eStatus				: E_Element_State_Long; // for HMI only as status
	
	fbPis				: FB_Piston;	
	
	//stPis_FillWater			: REFERENCE TO ST_Piston;
	//stPis_FillWaterDrain		: REFERENCE TO ST_Piston;
	//stPis_DrainTapWater		: REFERENCE TO ST_Piston;
	
	stPis_CWIn				: REFERENCE TO ST_Piston;
	stPis_CWOut				: REFERENCE TO ST_Piston;
	
	bTestingMode	:	BOOL	;//For testing purposes, to be deleted 
	bMoveStep		:	BOOL	;//For testing purposes, to be deleted 
	
	Call_TON	:	TON	;//Call ton for double request same object
	bTON_Active	:	BOOL	;
	
	// Temperature process control
	pc_TempCntrl	: REFERENCE TO FB_ProcessControl	;
	st_TempCntrl	: REFERENCE TO ST_ProcessControl	;
	bCntrlTemp		: BOOL	;
	bRunCIP			: BOOL	;
	
	ref_fbTankSensors			: REFERENCE TO FB_TankSensors;
	stTank_Level				: ST_Tank_Level;

	//888888888888888888888888888888888888888888
	stProdParam		: ST_Production_Parameter;
	//888888888888888888888888888888888888888888
	tonStirrer_time: TON;
	rTest: REAL := 16;
	bStirrerDirectionPositive: BOOL;
	
	delta_Tank_Volume		: REAL;
	memo_Tank_Level_start	: REAL;
	bRunOffline: BOOL;
	
	event_state_Update: INT;
	event_state_Update_sum: INT;
	event_state_Update_sum_last: INT;
	fbEvent_echo: FB_Event_echo;
	memo_Production_Storage_Mode: BOOL;
	memo_CIP_Pump_linked: BOOL;
	
	bStateUpdate_Available_HMI	: BOOL;

	
	
	fbFilling				: FB_Filling;		
	eFilling_State			: E_Filling_State;

END_VAR
VAR_IN_OUT

	fbTarget				: FB_Tank_Target;
	fbLineSource			: FB_Line_Source;
	fbLineTarget			: FB_Line_Target;
	fbTriBlenderSource		: FB_Line_Source;
	fbTriBlenderTarget		: FB_Line_Target;
	
	fbInterConnection_TriB	: FB_InterConnection;
	fbInterConnection_ProL	: FB_InterConnection;
	

	fb_PumpLine				: FB_Pump;
	fb_PumpTriBlender		: FB_Pump;
	fb_Stirrer				: FB_Pump;
END_VAR

act_GetReference();
act_Oper();
act_Call_Interface(); //There is no need to Call block if it comes from the outside
act_TempCntrl();
act_ExpirationTime();
act_Filling();

CASE eTank_Name OF
	E_Tank_Name.T1: sTank_Name:='Production Tank-T1';
	E_Tank_Name.T2: sTank_Name:='Production Tank-T2';
	E_Tank_Name.T3: sTank_Name:='Production Tank-T3';
	E_Tank_Name.T4: sTank_Name:='Production Tank-T4';
END_CASE

IF bTestingMode THEN;
	IF bMoveStep THEN;
		bMoveStep:=FALSE; 
	END_IF	
ELSE;
	bMoveStep:=TRUE; 
END_IF


IF stProdParam.bGetRecipe THEN;
	stProdParam.bGetRecipe:=FALSE;
	mGet_Recipe(indexRecipe:=stProdParam.hmiRecipeIndex+1);
END_IF
CASE eElementID	OF 
	E_Element_List.eTank_1,E_Element_List.eTank_2:;
		stProdParam.listRecipe:=g_Prod.listRecipe_Marinade;
	E_Element_List.eTank_3,E_Element_List.eTank_4:;
  		stProdParam.listRecipe:=g_Prod.listRecipe_Color;
END_CASE

stProdParam.timeRemainToStart:=mTimeRemainToStart();
stProdParam.timeProductionDuration:=mTimeProductionDuration();
refElement.ProdStatus:=stProdParam.eStatus;


IF refElement.m_Get_InterConnection()=E_InterConnection.NotConnected 
AND bReady
THEN;
	IF NOT bStateUpdate_Available_HMI THEN;
		refElement.fbEvent_echo.event();
		bStateUpdate_Available_HMI:=TRUE;
	END_IF	
ELSE; 
	IF bStateUpdate_Available_HMI THEN;
		refElement.fbEvent_echo.event();
		bStateUpdate_Available_HMI:=FALSE;
	END_IF
END_IF

m_Stirrer();
m_HMI();

ACTION _aCheck_Condition_Prod_End_active:
bStepDone:=FALSE;
IF fbInterConnection_ProL.bAvalableToDisconnect 
AND stProdParam.eStatus=E_Prod_Status.Active
THEN;
	bStepDone:=TRUE;
END_IF
END_ACTION

ACTION _aCheck_Condition_Product_active:
bStepDone:=FALSE;
IF fbInterConnection_ProL.bAvalableToConnect 
AND stProdParam.eStatus=E_Prod_Status.Active
THEN;
	bStepDone:=TRUE;
END_IF
END_ACTION

ACTION _aCheck_Condition_TriB_1_active_1:
bStepDone:=FALSE;
IF fbInterConnection_TriB.bAvalableToConnect
AND stProdParam.eStatus=E_Prod_Status.Active
AND m_Get_TriBlender_Clean()
THEN;
	bStepDone:=TRUE;
END_IF
END_ACTION

ACTION _aCheck_Condition_TriB_2_active:
bStepDone:=FALSE;
IF fbInterConnection_TriB.bAvalableToConnect 
AND stProdParam.eStatus=E_Prod_Status.Active
AND m_Get_TriBlender_Clean()
THEN;
	bStepDone:=TRUE;
END_IF
END_ACTION

ACTION _aClose_01_active:
bStepDone:=FALSE;
IF fbTarget.m_CheckStatus(eReqStatus:=E_Tank_Target.eClose) THEN;
	bStepDone:=TRUE;
END_IF
END_ACTION

ACTION _aClose_01_entry:
fbTarget.m_Run(eReqProc:=E_Tank_Target.eClose);
END_ACTION

ACTION _aClose_2_active:
bStepDone:=FALSE;
IF fbTarget.m_CheckStatus(eReqStatus:=E_Tank_Target.eClose) THEN;
	bStepDone:=TRUE;
END_IF
END_ACTION

ACTION _aClose_2_entry:
fbTarget.m_Run(eReqProc:=E_Tank_Target.eClose);
END_ACTION

ACTION _aClose_4_active:
bStepDone:=FALSE;
IF fbTarget.m_CheckStatus(eReqStatus:=E_Tank_Target.eClose) THEN;
	bStepDone:=TRUE;
END_IF
END_ACTION

ACTION _aClose_4_entry:
fbTarget.m_Run(eReqProc:=E_Tank_Target.eClose);
END_ACTION

ACTION _aClose_Drain_val_active:
//bStepDone:=FALSE;
IF fbTarget.m_CheckStatus(eReqStatus:=E_Tank_Target.eOpen) THEN;
(*ELSE
	fbTarget.m_Run(eReqProc:=E_Tank_Target.eOpen);*)
	bTON_Active:=TRUE;
END_IF
IF Call_TON.Q THEN
	bStepDone:=TRUE;
END_IF
END_ACTION

ACTION _aClose_Drain_val_entry:
bStepDone:=FALSE;
fbTarget.m_Run(eReqProc:=E_Tank_Target.eOpen);
bTON_Active:=FALSE;
END_ACTION

ACTION _aClose_Tank_active:
bStepDone:=FALSE;
IF fbTarget.m_CheckStatus(eReqStatus:=E_Tank_Target.eClose_DrainPipe) THEN;
	bStepDone:=TRUE;
END_IF
END_ACTION

ACTION _aClose_Tank_entry:
fbTarget.m_Run(eReqProc:=E_Tank_Target.eClose_DrainPipe);
END_ACTION

ACTION _aCollect_From_Prod_Line_active:
bStepDone:=FALSE;
delta_Tank_Volume:=ref_fbTankSensors.act_Volume-memo_Tank_Level_start;
IF FALSE 
OR delta_Tank_Volume>=stProdParam.stRecipe.Weight_to_Collect
OR Collect_From_Prod_Line.t>=T#40S
THEN;
	bStepDone:=TRUE;
END_IF
END_ACTION

ACTION _aCollect_From_TriB_Line_active:
bStepDone:=FALSE;
delta_Tank_Volume:=ref_fbTankSensors.act_Volume-memo_Tank_Level_start;
IF FALSE 
OR delta_Tank_Volume>=stProdParam.stRecipe.Weight_to_Collect
OR Collect_From_TriB_Line.t>=T#40S
THEN;
	bStepDone:=TRUE;
END_IF
END_ACTION

ACTION _aConn_Line_Source_TankA_active:
bStepDone:=FALSE;
IF fbLineSource.m_CheckStatus(eReqStatus:=E_Line_Source.eTank_A) THEN;
	bStepDone:=TRUE;
END_IF
END_ACTION

ACTION _aConn_Line_Source_TankA_entry:
fbLineSource.m_Run(eReqProc:=E_Line_Source.eTank_A);
END_ACTION

ACTION _aConn_Line_Source_TankB_active:
bStepDone:=FALSE;
IF fbLineSource.m_CheckStatus(eReqStatus:=E_Line_Source.eTank_B) THEN;
	bStepDone:=TRUE;
END_IF
END_ACTION

ACTION _aConn_Line_Source_TankB_entry:
fbLineSource.m_Run(eReqProc:=E_Line_Source.eTank_B);
END_ACTION

ACTION _aConn_Line_Target_TankA_active:
bStepDone:=FALSE;
IF fbLineTarget.m_CheckStatus(eReqStatus:=E_Line_Target.eTank_A) THEN;
	bTON_Active:=TRUE;
END_IF
IF Call_TON.Q THEN
	bStepDone:=TRUE;
END_IF
END_ACTION

ACTION _aConn_Line_Target_TankA_entry:
fbLineTarget.m_Run(eReqProc:=E_Line_Target.eTank_A);
bTON_Active:=FALSE;
END_ACTION

ACTION _aConn_Line_Target_TankB_active:
bStepDone:=FALSE;
IF fbLineTarget.m_CheckStatus(eReqStatus:=E_Line_Target.eTank_B) THEN;
	bTON_Active:=TRUE;
END_IF
IF Call_TON.Q THEN
	bStepDone:=TRUE;
END_IF
END_ACTION

ACTION _aConn_Line_Target_TankB_entry:
fbLineTarget.m_Run(eReqProc:=E_Line_Target.eTank_B);
bTON_Active:=FALSE;
END_ACTION

ACTION _aConn_Tank_active:
bStepDone:=FALSE;
IF fbTriBlenderSource.m_CheckStatus(eReqStatus:=E_Line_Source.eFillWater) 
//AND fbPis.m_CheckByRecipe(stPis:=stPis_FillWaterDrain, req:=E_Piston_Recipe_State.Release) 
THEN;
	bStepDone:=TRUE;
END_IF
END_ACTION

ACTION _aConn_Tank_entry:
fbTriBlenderSource.m_Run(eReqProc:=E_Line_Source.eFillWater);
//fbPis.m_SetByRecipe(stPis:=stPis_FillWaterDrain, req:=E_Piston_Recipe_State.Release);
END_ACTION

ACTION _aConn_Tri_Drain_active:
bStepDone:=FALSE;
IF fbTriBlenderTarget.m_CheckStatus(eReqStatus:=E_Line_Target.eDrain) THEN;
	bStepDone:=TRUE;
END_IF
END_ACTION

ACTION _aConn_Tri_Drain_entry:
fbTriBlenderTarget.m_Run(eReqProc:=E_Line_Target.eDrain);
END_ACTION

ACTION _aConn_Tri_TankA_2_active:
bStepDone:=FALSE;
IF fbTriBlenderSource.m_CheckStatus(eReqStatus:=E_Line_Source.eTank_A) THEN;
	bStepDone:=TRUE;
END_IF
END_ACTION

ACTION _aConn_Tri_TankA_2_entry:
fbTriBlenderSource.m_Run(eReqProc:=E_Line_Source.eTank_A);
END_ACTION

ACTION _aConn_Tri_TankB_2_active:
bStepDone:=FALSE;
IF fbTriBlenderSource.m_CheckStatus(eReqStatus:=E_Line_Source.eTank_B) THEN;
	bStepDone:=TRUE;
END_IF
END_ACTION

ACTION _aConn_Tri_TankB_2_entry:
fbTriBlenderSource.m_Run(eReqProc:=E_Line_Source.eTank_B);
END_ACTION

ACTION _aConn_Tri_TapWater_active:
bStepDone:=FALSE;
IF fbTriBlenderSource.m_CheckStatus(eReqStatus:=E_Line_Source.eTapWater) 
//AND fbPis.m_CheckByRecipe(stPis:=stPis_DrainTapWater, req:=E_Piston_Recipe_State.Release) 
THEN;
	bTON_Active:=TRUE;
END_IF
IF Call_TON.Q THEN
	bStepDone:=TRUE;
END_IF
END_ACTION

ACTION _aConn_Tri_TapWater_entry:
fbTriBlenderSource.m_Run(eReqProc:=E_Line_Source.eTapWater);
//fbPis.m_SetByRecipe(stPis:=stPis_DrainTapWater, req:=E_Piston_Recipe_State.Release);
bTON_Active:=FALSE;
END_ACTION

ACTION _aConn_Tri_ToTankA_1_active:
bStepDone:=FALSE;
IF fbTriBlenderTarget.m_CheckStatus(eReqStatus:=E_Line_Target.eTank_A) THEN;
	bStepDone:=TRUE;
END_IF
END_ACTION

ACTION _aConn_Tri_ToTankA_1_entry:
fbTriBlenderTarget.m_Run(eReqProc:=E_Line_Target.eTank_A);
END_ACTION

ACTION _aConn_Tri_ToTankA_2_active:
bStepDone:=FALSE;
IF fbTriBlenderTarget.m_CheckStatus(eReqStatus:=E_Line_Target.eTank_A) THEN;
	bStepDone:=TRUE;
END_IF
END_ACTION

ACTION _aConn_Tri_ToTankA_2_entry:
fbTriBlenderTarget.m_Run(eReqProc:=E_Line_Target.eTank_A);
END_ACTION

ACTION _aConn_Tri_ToTankB_1_active:
bStepDone:=FALSE;
IF fbTriBlenderTarget.m_CheckStatus(eReqStatus:=E_Line_Target.eTank_B) THEN;
	bStepDone:=TRUE;
END_IF
END_ACTION

ACTION _aConn_Tri_ToTankB_1_entry:
fbTriBlenderTarget.m_Run(eReqProc:=E_Line_Target.eTank_B);
END_ACTION

ACTION _aConn_Tri_ToTankB_2_active:
bStepDone:=FALSE;
IF fbTriBlenderTarget.m_CheckStatus(eReqStatus:=E_Line_Target.eTank_B) THEN;
	bStepDone:=TRUE;
END_IF
END_ACTION

ACTION _aConn_Tri_ToTankB_2_entry:
fbTriBlenderTarget.m_Run(eReqProc:=E_Line_Target.eTank_B);
END_ACTION

ACTION _aConn_TriB_Color_active_1:
bStepDone:=FALSE;
IF fbTriBlender_Select.m_CheckStatus(eReqStatus:=E_TriBlenderSelect.eColor) THEN;
	bStepDone:=TRUE;
END_IF
END_ACTION

ACTION _aConn_TriB_Color_entry_1:
fbTriBlender_Select.m_Set_Request(eSetReg:=E_TriBlenderSelect.eColor);
END_ACTION

ACTION _aConn_TriB_Marinade_active_1:
bStepDone:=FALSE;
IF fbTriBlender_Select.m_CheckStatus(eReqStatus:=E_TriBlenderSelect.eMarinade) THEN;
	bStepDone:=TRUE;
END_IF
END_ACTION

ACTION _aConn_TriB_Marinade_entry_1:
fbTriBlender_Select.m_Set_Request(eSetReg:=E_TriBlenderSelect.eMarinade);
END_ACTION

ACTION _aDis_Conn_Tank_active:
bStepDone:=FALSE;
IF fbTriBlenderSource.m_CheckStatus(eReqStatus:=E_Line_Source.eClose) 
AND fbTriBlenderTarget.m_CheckStatus(eReqStatus:=E_Line_Target.eDrain) 
THEN;
	bStepDone:=TRUE;
END_IF
END_ACTION

ACTION _aDis_Conn_Tank_entry:
fbTriBlenderSource.m_Run(eReqProc:=E_Line_Source.eClose);
fbTriBlenderTarget.m_Run(eReqProc:=E_Line_Target.eDrain);
END_ACTION

ACTION _aDisconn_Tri_Tank_active:
bStepDone:=FALSE;
IF fbTriBlenderSource.m_CheckStatus(eReqStatus:=E_Line_Source.eClose) THEN;
	bTON_Active:=TRUE;
END_IF
IF Call_TON.Q THEN
	bStepDone:=TRUE;
END_IF
END_ACTION

ACTION _aDisconn_Tri_Tank_entry:
fbTriBlenderSource.m_Run(eReqProc:=E_Line_Source.eClose);
bTON_Active:=FALSE;
END_ACTION

ACTION _aDisconnect_TapWater_02_active:
bStepDone:=FALSE;
IF fbTriBlenderSource.m_CheckStatus(eReqStatus:=E_Line_Source.eDrain) THEN;
	bStepDone:=TRUE;
END_IF
END_ACTION

ACTION _aDisconnect_TapWater_02_entry:
fbTriBlenderSource.m_Run(eReqProc:=E_Line_Source.eDrain);
END_ACTION

ACTION _aDissolving_entry:
bDisolvingProcess_Done:=FALSE;
bDisolvingProcess_Active:=FALSE;
END_ACTION

ACTION _aDissolving_Proc_active:
bStepDone:=FALSE;

IF bDisolvingProcess_Done 
//AND fbDissolving.bD
THEN;
	
END_IF
END_ACTION

ACTION _aDissolving_Proc_entry:

bDisolvingProcess_Active:=TRUE;
fbDissolving.mRun();
END_ACTION

ACTION _aDissolving_Proc_exit:
bDisolvingProcess_Done:=FALSE;
bDisolvingProcess_Active:=FALSE;
END_ACTION

ACTION _aDone_entry:
eProcess:=E_Element_Process.eNone;
eReq:=E_Request_List.eNone;
bRun:=FALSE;
bDone:=TRUE;
END_ACTION

ACTION _aDrain_All_Marinade_Lines_active:
bStepDone:=FALSE;
IF TRUE
//AND fbTarget.m_CheckStatus(eReqStatus:=E_Tank_Target.eClose_DrainPipe) 
AND fbTriBlenderSource.m_CheckStatus(eReqStatus:=E_Line_Source.eDrain)
AND fbTriBlenderTarget.m_CheckStatus(eReqStatus:=E_Line_Target.eDrain)
AND fbTriBlender_Select.m_CheckStatus(eReqStatus:=E_TriBlenderSelect.eDrain)
AND TRUE
AND TRUE
THEN;
	bStepDone:=TRUE;
END_IF
END_ACTION

ACTION _aDrain_All_Marinade_Lines_entry:
//fbTarget.m_Run(eReqProc:=E_Tank_Target.eClose_DrainPipe);
fbTriBlenderSource.m_Run(eReqProc:=E_Line_Source.eDrain);
fbTriBlenderTarget.m_Run(eReqProc:=E_Line_Target.eDrain);
fbTriBlender_Select.m_Set_Request(eSetReg:=E_TriBlenderSelect.eDrain);
END_ACTION

ACTION _aDrain_Pipe_active:
bStepDone:=FALSE;
IF fbTarget.m_CheckStatus(eReqStatus:=E_Tank_Target.eClose_DrainPipe) THEN;
	bTON_Active:=TRUE;
END_IF
IF Call_TON.Q THEN
	bStepDone:=TRUE;
END_IF
END_ACTION

ACTION _aDrain_Pipe_Close_active:
bStepDone:=FALSE;
IF fbTarget.m_CheckStatus(eReqStatus:=E_Tank_Target.eClose) THEN;
	bStepDone:=TRUE;
END_IF
END_ACTION

ACTION _aDrain_Pipe_Close_entry:
fbTarget.m_Run(eReqProc:=E_Tank_Target.eClose);
END_ACTION

ACTION _aDrain_Pipe_entry:
fbTarget.m_Run(eReqProc:=E_Tank_Target.eClose_DrainPipe);
bTON_Active:=FALSE;
END_ACTION

ACTION _aDrain_Production_Line_active:
bStepDone:=FALSE;
IF TRUE
AND fbTarget.m_CheckStatus(eReqStatus:=E_Tank_Target.eClose_DrainPipe) 
AND fbLineSource.m_CheckStatus(eReqStatus:=E_Line_Source.eDrain)
AND fbLineTarget.m_CheckStatus(eReqStatus:=E_Line_Target.eDrain)
AND TRUE
THEN;
	bStepDone:=TRUE;
END_IF
END_ACTION

ACTION _aDrain_Production_Line_entry:
fbTarget.m_Run(eReqProc:=E_Tank_Target.eClose_DrainPipe);
fbLineSource.m_Run(eReqProc:=E_Line_Source.eDrain);
fbLineTarget.m_Run(eReqProc:=E_Line_Target.eDrain);
END_ACTION

ACTION _aDrain_Tri_Line_active:
bStepDone:=FALSE;
IF fbTriBlenderTarget.m_CheckStatus(eReqStatus:=E_Line_Target.eDrain) THEN;
	bStepDone:=TRUE;
END_IF
END_ACTION

ACTION _aDrain_Tri_Line_entry:
fbTriBlenderTarget.m_Run(eReqProc:=E_Line_Target.eDrain);
END_ACTION

ACTION _aDrain_Tri_ToDrain_active:
bStepDone:=FALSE;
IF fbTriBlenderTarget.m_CheckStatus(eReqStatus:=E_Line_Target.eDrain) THEN;
	bTON_Active:=TRUE;
END_IF
IF Call_TON.Q THEN
	bStepDone:=TRUE;
END_IF

(*
delta_Tank_Volume:=ref_fbTankSensors.act_Volume-memo_Tank_Level_start;
IF bStepDone
AND  
AND (delta_Tank_Volume>=stProdParam.stRecipe.Weight_to_Drain
	OR Drain_Tri_ToDrain.t>=T#30S)
THEN;
	//bStepDone:=TRUE;
ELSE;
	bStepDone:=FALSE;
END_IF
*)
END_ACTION

ACTION _aDrain_Tri_ToDrain_entry:
fbTriBlenderTarget.m_Run(eReqProc:=E_Line_Target.eDrain);
bTON_Active:=FALSE;
END_ACTION

ACTION _aDrain_Tri_ToTankA_active:
bStepDone:=FALSE;
IF fbTriBlenderTarget.m_CheckStatus(eReqStatus:=E_Line_Target.eTank_A) THEN;
	bTON_Active:=TRUE;
END_IF
IF Call_TON.Q THEN
	bStepDone:=TRUE;
END_IF
END_ACTION

ACTION _aDrain_Tri_ToTankA_entry:
fbTriBlenderTarget.m_Run(eReqProc:=E_Line_Target.eTank_A);
bTON_Active:=FALSE;
END_ACTION

ACTION _aDrain_Tri_ToTankB_active:
bStepDone:=FALSE;
IF fbTriBlenderTarget.m_CheckStatus(eReqStatus:=E_Line_Target.eTank_B) THEN;
	bTON_Active:=TRUE;
END_IF
IF Call_TON.Q THEN
	bStepDone:=TRUE;
END_IF
END_ACTION

ACTION _aDrain_Tri_ToTankB_entry:
fbTriBlenderTarget.m_Run(eReqProc:=E_Line_Target.eTank_B);
bTON_Active:=FALSE;
END_ACTION

ACTION _aDrain_Trib_Line_01_active:
bStepDone:=FALSE;
IF fbTriBlender_Select.m_CheckStatus(eReqStatus:=E_TriBlenderSelect.eDrain) THEN;
	bStepDone:=TRUE;
END_IF
END_ACTION

ACTION _aDrain_Trib_Line_01_entry:
fbTriBlender_Select.m_Set_Request(eSetReg:=E_TriBlenderSelect.eDrain);
END_ACTION

ACTION _aDrain_Trib_Line_02_active:
bStepDone:=FALSE;
IF fbTriBlender_Select.m_CheckStatus(eReqStatus:=E_TriBlenderSelect.eDrain)
OR fbTriBlender_Select.m_CheckStatus(eReqStatus:=E_TriBlenderSelect.eMarinade) THEN;//marinade =>> drain time finish
	bStepDone:=TRUE;
END_IF
END_ACTION

ACTION _aDrain_Trib_Line_02_entry:
fbTriBlender_Select.m_Set_Request(eSetReg:=E_TriBlenderSelect.eDrain);
END_ACTION

ACTION _aDraining_Time_active:
bStepDone:=FALSE;
IF stTank_Level.e_state=E_Tank_Level.eEmpty THEN;
	bStepDone:=TRUE;
END_IF
END_ACTION

ACTION _aDrainOpen_01_active:
bStepDone:=FALSE;
IF fbTarget.m_CheckStatus(eReqStatus:=E_Tank_Target.eDrain) THEN;
	bStepDone:=TRUE;
END_IF
END_ACTION

ACTION _aDrainOpen_01_entry:
fbTarget.m_Run(eReqProc:=E_Tank_Target.eDrain);
END_ACTION

ACTION _aDriin_Tank_active:
bStepDone:=FALSE;
IF stTank_Level.e_state=E_Tank_Level.eEmpty THEN;
	bStepDone:=TRUE;
END_IF
END_ACTION

ACTION _aDriin_Tank_entry:
fbTarget.m_Run(eReqProc:=E_Tank_Target.eDrain);
END_ACTION

ACTION _aInit_Base_active:
bStepDone:=FALSE;
IF TRUE
AND refState_Long<>E_Element_State_Long.eProduction
AND fbTarget.m_CheckStatus(eReqStatus:=E_Tank_Target.eClose_DrainPipe) 
AND TRUE
THEN;
	bStepDone:=TRUE;
ELSIF refState_Long=E_Element_State_Long.eProduction THEN;
	bStepDone:=TRUE;
END_IF
END_ACTION

ACTION _aInit_Base_entry:
IF refState_Long<>E_Element_State_Long.eProduction THEN;	
	fb_PumpLine.m_Stop();
	fbTarget.m_Run(eReqProc:=E_Tank_Target.eClose_DrainPipe);
END_IF
END_ACTION

ACTION _aInit_Production_Line_active:
bStepDone:=FALSE;
IF TRUE
AND refState_Long<>E_Element_State_Long.eProduction
AND fbTarget.m_CheckStatus(eReqStatus:=E_Tank_Target.eClose_DrainPipe) 
AND fbLineSource.m_CheckStatus(eReqStatus:=E_Line_Source.eDrain)
AND fbLineTarget.m_CheckStatus(eReqStatus:=E_Line_Target.eDrain)
AND (NOT fbInterConnection_ProL.bActive)
AND TRUE
THEN;
	bStepDone:=TRUE;
ELSIF refState_Long=E_Element_State_Long.eProduction THEN;
	bStepDone:=TRUE;
END_IF
END_ACTION

ACTION _aInit_Production_Line_entry:
IF refState_Long<>E_Element_State_Long.eProduction THEN;	
	fb_PumpLine.m_Stop();
	fbTarget.m_Run(eReqProc:=E_Tank_Target.eClose_DrainPipe);
	fbLineSource.m_Run(eReqProc:=E_Line_Source.eDrain);
	fbLineTarget.m_Run(eReqProc:=E_Line_Target.eDrain);
	fbInterConnection_ProL.reqDisconnect:=TRUE;
END_IF
END_ACTION

ACTION _aInit_Tank_active:
SFCReset:=FALSE;
END_ACTION

ACTION _aInit_Tank_exit:
IF eProcess=E_Element_Process.eFill_Water THEN;
	mClearProduction(state:=E_Element_State_Long.eOff);
END_IF

eProcess:=E_Element_Process.eNone;
eReq:=E_Request_List.eNone;
memo_Production_Storage_Mode:=FALSE;
END_ACTION

ACTION _aInit_TriBlender_Line_active:
bStepDone:=FALSE;
IF TRUE
AND fbTarget.m_CheckStatus(eReqStatus:=E_Tank_Target.eClose_DrainPipe) 
AND fbTriBlenderSource.m_CheckStatus(eReqStatus:=E_Line_Source.eDrain)
AND fbTriBlenderTarget.m_CheckStatus(eReqStatus:=E_Line_Target.eDrain)
AND fbTriBlender_Select.m_CheckStatus(eReqStatus:=E_TriBlenderSelect.eDrain)
AND (NOT fbInterConnection_TriB.bActive)
AND TRUE
THEN;
	bStepDone:=TRUE;
END_IF
END_ACTION

ACTION _aInit_TriBlender_Line_entry:
fb_PumpTriBlender.m_Stop();
fbTarget.m_Run(eReqProc:=E_Tank_Target.eClose_DrainPipe);
fbTriBlenderSource.m_Run(eReqProc:=E_Line_Source.eDrain);
fbTriBlenderTarget.m_Run(eReqProc:=E_Line_Target.eDrain);
fbTriBlender_Select.m_Set_Request(eSetReg:=E_TriBlenderSelect.eDrain);
fbInterConnection_TriB.reqDisconnect:=TRUE;
fbDissolving.mResetCycle();
END_ACTION

ACTION _aInterConnect_Prod_active:
bStepDone:=FALSE;
IF fbInterConnection_ProL.bActive THEN;
	bStepDone:=TRUE;
END_IF
END_ACTION

ACTION _aInterConnect_Prod_Dis_active:
bStepDone:=FALSE;
IF NOT fbInterConnection_ProL.bActive THEN;
	bStepDone:=TRUE;
END_IF
END_ACTION

ACTION _aInterConnect_Prod_Dis_entry:
fbInterConnection_ProL.reqDisconnect:=TRUE;
END_ACTION

ACTION _aInterConnect_Prod_entry:
fbInterConnection_ProL.reqConnect:=TRUE;

IF trn_Tank_Marinade THEN;
	//fbElement[E_Element_List.eTriBlender_Marinada].m_Set_Dissolveng_active_memo();
ELSIF trn_Tank_Color THEN;
	//fbElement[E_Element_List.eTriBlender_Color].m_Set_Dissolveng_active_memo();
END_IF
END_ACTION

ACTION _aInterConnect_TriB_1_active:
bStepDone:=FALSE;
IF fbInterConnection_TriB.bActive THEN;
	bStepDone:=TRUE;
END_IF
END_ACTION

ACTION _aInterConnect_TriB_1_entry:
fbInterConnection_TriB.reqConnect:=TRUE;
END_ACTION

ACTION _aInterConnect_TriB_2_active:
bStepDone:=FALSE;
IF fbInterConnection_TriB.bActive THEN;
	bStepDone:=TRUE;
	
	refElement.m_Set_Dissolveng_active_memo();
	IF trn_Tank_Marinade THEN;
		fbElement[E_Element_List.eTriBlender_Marinada].m_Set_Dissolveng_active_memo();
	ELSIF trn_Tank_Color THEN;
		fbElement[E_Element_List.eTriBlender_Color].m_Set_Dissolveng_active_memo();
	ELSE;
		bStepDone:=FALSE;
	END_IF	
	
END_IF
END_ACTION

ACTION _aInterConnect_TriB_2_entry:
fbInterConnection_TriB.reqConnect:=TRUE;
END_ACTION

ACTION _aInterConnect_TriB_Dis_1_active:
bStepDone:=FALSE;
IF NOT fbInterConnection_TriB.bActive THEN;
	bStepDone:=TRUE;
END_IF
END_ACTION

ACTION _aInterConnect_TriB_Dis_1_entry:
fbInterConnection_TriB.reqDisconnect:=TRUE;
END_ACTION

ACTION _aInterConnect_TriB_Dis_2_active:
bStepDone:=FALSE;
IF NOT fbInterConnection_TriB.bActive THEN;
	bStepDone:=TRUE;
END_IF
END_ACTION

ACTION _aInterConnect_TriB_Dis_2_entry:
fbInterConnection_TriB.reqDisconnect:=TRUE;
END_ACTION

ACTION _aLineSource_Close_active:
bStepDone:=FALSE;
IF fbLineSource.m_CheckStatus(eReqStatus:=E_Line_Source.eClose) 
THEN;
	bStepDone:=TRUE;
END_IF
END_ACTION

ACTION _aLineSource_Close_entry:
fbLineSource.m_Run(eReqProc:=E_Line_Source.eClose);
END_ACTION

ACTION _aLineSource_TapWater_active:
bStepDone:=FALSE;
IF fbLineSource.m_CheckStatus(eReqStatus:=E_Line_Source.eTapWater) 
THEN;
	bStepDone:=TRUE;
END_IF
END_ACTION

ACTION _aLineSource_TapWater_entry:
fbLineSource.m_Run(eReqProc:=E_Line_Source.eTapWater);
bTON_Active:=FALSE;
END_ACTION

ACTION _aLineTarget_Drain_1_active:
bStepDone:=FALSE;
IF fbLineTarget.m_CheckStatus(eReqStatus:=E_Line_Target.eDrain) THEN;
	bStepDone:=TRUE;
END_IF
END_ACTION

ACTION _aLineTarget_Drain_1_entry:
fbLineTarget.m_Run(eReqProc:=E_Line_Target.eDrain);
END_ACTION

ACTION _aLineTarget_Drain_2_active:
bStepDone:=FALSE;
IF fbLineTarget.m_CheckStatus(eReqStatus:=E_Line_Target.eDrain) THEN;
	bTON_Active:=TRUE;
END_IF
IF Call_TON.Q THEN
	bStepDone:=TRUE;
END_IF
END_ACTION

ACTION _aLineTarget_Drain_2_entry:
fbLineTarget.m_Run(eReqProc:=E_Line_Target.eDrain);
bTON_Active:=FALSE;
END_ACTION

ACTION _aLineTarget_TankA_active:
bStepDone:=FALSE;
IF fbLineTarget.m_CheckStatus(eReqStatus:=E_Line_Target.eTank_A) THEN;
	bTON_Active:=TRUE;
END_IF
IF Call_TON.Q THEN
	bStepDone:=TRUE;
END_IF
END_ACTION

ACTION _aLineTarget_TankA_entry:
fbLineTarget.m_Run(eReqProc:=E_Line_Target.eTank_A);
bTON_Active:=FALSE;
END_ACTION

ACTION _aLineTarget_TankB_active:
bStepDone:=FALSE;
IF fbLineTarget.m_CheckStatus(eReqStatus:=E_Line_Target.eTank_B) THEN;
	bTON_Active:=TRUE;
END_IF
IF Call_TON.Q THEN
	bStepDone:=TRUE;
END_IF
END_ACTION

ACTION _aLineTarget_TankB_entry:
fbLineTarget.m_Run(eReqProc:=E_Line_Target.eTank_B);
bTON_Active:=FALSE;
END_ACTION

ACTION _aOpen_Drain_Pipe_active:
bStepDone:=FALSE;
IF fbTarget.m_CheckStatus(eReqStatus:=E_Tank_Target.eClose_DrainPipe) THEN;
	bStepDone:=TRUE;
END_IF
END_ACTION

ACTION _aOpen_Drain_Pipe_entry:
fbTarget.m_Run(eReqProc:=E_Tank_Target.eClose_DrainPipe);
END_ACTION

ACTION _aPumpLine_Auto_1_entry:
//fb_PumpLine.m_Auto();
END_ACTION

ACTION _aPumpLine_Start_1_active:

END_ACTION

ACTION _aPumpLine_Start_1_entry:
fb_PumpLine.m_Run(RPM:=stProdParam.stRecipe.FlowRate_Production);
END_ACTION

ACTION _aPumpLine_Start_2_entry:
fb_PumpLine.m_Run(RPM:=stProdParam.stRecipe.FlowRate_Production);
memo_Tank_Level_start:=ref_fbTankSensors.act_Volume;
END_ACTION

ACTION _aPumpLine_Stop_1_entry:
fb_PumpLine.m_Stop();
END_ACTION

ACTION _aPumpLine_Stop_2_entry:

IF trn_Tank_Marinade THEN;
	fb_PumpLine.m_Stop();
END_IF
END_ACTION

ACTION _aPumpLine_Stop_3_entry:
fb_PumpLine.m_Stop();
END_ACTION

ACTION _aPumpLine_Stop_4_entry:
fb_PumpLine.m_Stop();
END_ACTION

ACTION _aReady_active:


CASE refElement.eState_Long OF
	E_Element_State_Long.eOff,E_Element_State_Long.eStandby:;
			IF eReq=E_Request_List.eDrain THEN;
				eProcess:=E_Element_Process.eDrain;
			END_IF

	E_Element_State_Long.eCIP_5_Done:;
			IF eReq=E_Request_List.eWaterPrepare THEN;
				eProcess:=E_Element_Process.eFill_Water;
			END_IF	
			
